// TwinCAT 3 PLC project Syn_Config
// Title: SynConfig
// Company: Syntegon Group
// ProjectVersion: 2.4.0.0
// Description: Parameter sets the RPP configurator writes and the application takes over (ADR 0017).
// ProgramVersion: 3.1.4026.28
// libraries:
//   Tc2_Standard,newest,Beckhoff Automation GmbH
//   SynVisu, * (Syntegon Group)
// project tree:
//   DUTs/ E_ConfigCommand.TcDUT, E_ConfigCommandResult.TcDUT, E_ConfigFieldType.TcDUT, E_ConfigResult.TcDUT, ST_ConfigBodyComponent.TcDUT, ST_ConfigBodyComponentParam.TcDUT, ST_ConfigBodyComponentSet.TcDUT, ST_ConfigCartesian.TcDUT, ST_ConfigCartesianParam.TcDUT, ST_ConfigCartesianSet.TcDUT, ST_ConfigCommand.TcDUT, ST_ConfigCommandStatus.TcDUT, ST_ConfigConveyor.TcDUT, ST_ConfigConveyorParam.TcDUT, ST_ConfigConveyorSet.TcDUT, ST_ConfigDelta.TcDUT, ST_ConfigDeltaParam.TcDUT, ST_ConfigDeltaSet.TcDUT, ST_ConfigMachine.TcDUT, ST_ConfigManifest.TcDUT, ST_ConfigManifestEntry.TcDUT, ST_ConfigRecipeField.TcDUT, ST_ConfigRecipeSet.TcDUT, ST_ConfigStaging.TcDUT, ST_ConfigStatus.TcDUT, ST_ConfigTopology.TcDUT, ST_ConfigTopologyKind.TcDUT, ST_ConfigTopologyLink.TcDUT, ST_ConfigTopologyLinks.TcDUT, ST_ConfigTopologyNode.TcDUT, ST_ConfigTopologyRole.TcDUT, ST_ConfigXtsGantry.TcDUT, ST_ConfigXtsGantryParam.TcDUT, ST_ConfigXtsGantrySet.TcDUT, ST_ConfigXtsLoop.TcDUT, ST_ConfigXtsLoopParam.TcDUT, ST_ConfigXtsLoopSet.TcDUT
//   GVLs/ CONFIG_GlobalConst.TcGVL, CONFIG_GlobalConst_Param.TcGVL
//   POUs/ _FB_ConfigBodyComponent.TcPOU, _FB_ConfigCartesian.TcPOU, _FB_ConfigComponent.TcPOU, _FB_ConfigConveyor.TcPOU, _FB_ConfigDelta.TcPOU, _FB_ConfigMachine.TcPOU, _FB_ConfigSensor.TcPOU, _FB_ConfigStation.TcPOU, _FB_ConfigTopology.TcPOU, _FB_ConfigVision.TcPOU, _FB_ConfigXtsGantry.TcPOU, _FB_ConfigXtsLoop.TcPOU, _FC_GetVersionSynConfig.TcPOU
// (motion and I/O tree: see PLC project syn_visu)
// real-time tasks:
//   TASK PlcTask: cycle T#10ms, priority 20, ADS port 350
//   TASK TestTask: cycle T#10ms, priority 21, ADS port 351

// ---- DUTs/E_ConfigCommand.TcDUT
{attribute 'qualified_only'}
{attribute 'strict'}
TYPE E_ConfigCommand :
(
	(* What a machine command asks the application (config protocol 3). Values are part of the gateway contract:
	   append, never renumber. *)
	NONE := 0,
	START := 1,
	STOP := 2,
	RESET := 3
) UINT;
END_TYPE

// ---- DUTs/E_ConfigCommandResult.TcDUT
{attribute 'qualified_only'}
{attribute 'strict'}
TYPE E_ConfigCommandResult :
(
	(* What the application made of the last machine command. Values are part of the gateway contract: append, never
	   renumber. *)
	NONE := 0,		// nothing asked since the PLC started
	ACCEPTED := 1,
	REJECTED := 2	// ST_ConfigCommandStatus.sMessage says why
) UINT;
END_TYPE

// ---- DUTs/E_ConfigFieldType.TcDUT
{attribute 'qualified_only'}
{attribute 'strict'}
TYPE E_ConfigFieldType :
(
	(* How a recipe field's value is kept (config protocol 3). Every value travels as LREAL. Values are part of the
	   gateway contract: append, never renumber. *)
	NUMBER := 0,	// any number within fMin..fMax
	INTEGER := 1,	// a whole number within fMin..fMax, e.g. picks per cycle
	SWITCH := 2,	// on or off: 1 or 0
	CHOICE := 3		// one of the named choices: 0..nChoiceCount-1
) UINT;
END_TYPE

// ---- DUTs/E_ConfigResult.TcDUT
{attribute 'qualified_only'}
{attribute 'strict'}
TYPE E_ConfigResult :
(
	(* What became of the last staged parameter set. Values are part of the gateway contract: append, never renumber. *)
	NONE := 0,		// nothing staged since the PLC started
	PENDING := 1,	// staged, waiting for the application to allow taking it over
	APPLIED := 2,	// taken over (or reset to the program values)
	REJECTED := 3	// not taken over; ST_ConfigStatus.sMessage says why
) UINT;
END_TYPE

// ---- DUTs/ST_ConfigBodyComponent.TcDUT
TYPE ST_ConfigBodyComponent :
STRUCT
	(* vo_Config of _FB_ConfigVision, _FB_ConfigSensor and _FB_ConfigStation: the gateway writes stStaging and
	   stStaged, reads stStatus and stActive. *)
	stStaging : ST_ConfigStaging;
	stStaged : ST_ConfigBodyComponentParam;
	stStatus : ST_ConfigStatus;
	stActive : ST_ConfigBodyComponentParam; // effective values: the active set while one is valid, else the program values
END_STRUCT
END_TYPE

// ---- DUTs/ST_ConfigBodyComponentParam.TcDUT
TYPE ST_ConfigBodyComponentParam :
STRUCT
	(* The parameter set of a component drawn from its bodies (vision system, product sensor, station): what the
	   configurator writes, never its bodies (hardware). Members as in SynVisu.ST_VisuDetectorConfig. *)
	stPose : SynVisu.ST_VisuPose; // MCS
	stOriginShift : SynVisu.ST_VisuPosition; // mm in the component's local frame
	nZoneCount : UINT;
	aZones : ARRAY[0..SynVisu.VISU_GlobalConst_Param.VISU_un_MAX_ZONES - 1] OF SynVisu.ST_VisuZone;
END_STRUCT
END_TYPE

// ---- DUTs/ST_ConfigBodyComponentSet.TcDUT
TYPE ST_ConfigBodyComponentSet :
STRUCT
	(* The active parameter set of a vision system, product sensor or station as the application keeps it, in a
	   VAR PERSISTENT variable passed to m_Cycle of _FB_ConfigVision, _FB_ConfigSensor or _FB_ConfigStation. *)
	bValid : BOOL; // FALSE: no set active, the program values apply
	nVersion : UDINT; // version of stParam
	nLastVersion : UDINT; // last version handed out; versions never repeat, also after a reset
	stParam : ST_ConfigBodyComponentParam;
END_STRUCT
END_TYPE

// ---- DUTs/ST_ConfigCartesian.TcDUT
TYPE ST_ConfigCartesian :
STRUCT
	(* vo_Config of _FB_ConfigCartesian: the gateway writes stStaging and stStaged, reads stStatus and stActive. *)
	stStaging : ST_ConfigStaging;
	stStaged : ST_ConfigCartesianParam;
	stStatus : ST_ConfigStatus;
	stActive : ST_ConfigCartesianParam; // effective values: the active set while one is valid, else the program values
END_STRUCT
END_TYPE

// ---- DUTs/ST_ConfigCartesianParam.TcDUT
TYPE ST_ConfigCartesianParam :
STRUCT
	(* A Cartesian robot's parameter set: what the configurator writes, never its axes, strokes or rail height
	   (hardware). Members as in SynVisu.ST_VisuCartesianConfig. *)
	stPose : SynVisu.ST_VisuPose; // MCS, axis origin X = Y = 0 with Z up
	stOriginShift : SynVisu.ST_VisuPosition; // mm in the robot's local frame
	nZoneCount : UINT;
	aZones : ARRAY[0..SynVisu.VISU_GlobalConst_Param.VISU_un_MAX_ZONES - 1] OF SynVisu.ST_VisuZone;
	nFingerCount : UINT; // gripper fingers with their flange offsets (config protocol 2, ADR 0018)
	aFingers : ARRAY[0..SynVisu.VISU_GlobalConst_Param.VISU_un_MAX_FINGERS - 1] OF SynVisu.ST_VisuFinger;
	stLimitArea : SynVisu.ST_VisuLimitArea; // bActive = FALSE: none
	stTcpLimitArea : SynVisu.ST_VisuLimitArea; // bActive = FALSE: none
END_STRUCT
END_TYPE

// ---- DUTs/ST_ConfigCartesianSet.TcDUT
TYPE ST_ConfigCartesianSet :
STRUCT
	(* A Cartesian robot's active parameter set as the application keeps it, in a VAR PERSISTENT variable passed to
	   _FB_ConfigCartesian.m_Cycle. *)
	bValid : BOOL; // FALSE: no set active, the program values apply
	nVersion : UDINT; // version of stParam
	nLastVersion : UDINT; // last version handed out; versions never repeat, also after a reset
	stParam : ST_ConfigCartesianParam;
END_STRUCT
END_TYPE

// ---- DUTs/ST_ConfigCommand.TcDUT
TYPE ST_ConfigCommand :
STRUCT
	(* A machine command, written by the gateway with bRequested last (config protocol 3). The machine FB clears
	   bRequested once the application answered it. *)
	nCommandId : UDINT; // chosen by the gateway; ST_ConfigCommandStatus.nHandledCommandId names it once answered
	eCommand : E_ConfigCommand;
	bRequested : BOOL; // TRUE: the command waits for the application's answer
END_STRUCT
END_TYPE

// ---- DUTs/ST_ConfigCommandStatus.TcDUT
TYPE ST_ConfigCommandStatus :
STRUCT
	nHandledCommandId : UDINT; // nCommandId of the last command the application answered
	eResult : E_ConfigCommandResult; // what the application made of it
	sMessage : STRING(80); // why it was rejected; empty otherwise
END_STRUCT
END_TYPE

// ---- DUTs/ST_ConfigConveyor.TcDUT
TYPE ST_ConfigConveyor :
STRUCT
	(* vo_Config of _FB_ConfigConveyor: the gateway writes stStaging and stStaged, reads stStatus and stActive. *)
	stStaging : ST_ConfigStaging;
	stStaged : ST_ConfigConveyorParam;
	stStatus : ST_ConfigStatus;
	stActive : ST_ConfigConveyorParam; // effective values: the active set while one is valid, else the program values
END_STRUCT
END_TYPE

// ---- DUTs/ST_ConfigConveyorParam.TcDUT
TYPE ST_ConfigConveyorParam :
STRUCT
	(* A conveyor's parameter set: what the configurator writes, never the belt's length or width (hardware).
	   Members as in SynVisu.ST_VisuConveyorConfig. *)
	stPose : SynVisu.ST_VisuPose; // MCS, belt start on the belt surface; local +X = conveying direction
	stOriginShift : SynVisu.ST_VisuPosition; // mm in the local frame from stPose: origin of the belt coordinates
	nProductTypeCount : UINT;
	aProductTypes : ARRAY[0..SynVisu.VISU_GlobalConst_Param.VISU_un_MAX_PRODUCT_TYPES - 1] OF SynVisu.ST_VisuProductType;
END_STRUCT
END_TYPE

// ---- DUTs/ST_ConfigConveyorSet.TcDUT
TYPE ST_ConfigConveyorSet :
STRUCT
	(* A conveyor's active parameter set as the application keeps it, in a VAR PERSISTENT variable passed to
	   _FB_ConfigConveyor.m_Cycle. *)
	bValid : BOOL; // FALSE: no set active, the program values apply
	nVersion : UDINT; // version of stParam
	nLastVersion : UDINT; // last version handed out; versions never repeat, also after a reset
	stParam : ST_ConfigConveyorParam;
END_STRUCT
END_TYPE

// ---- DUTs/ST_ConfigDelta.TcDUT
TYPE ST_ConfigDelta :
STRUCT
	(* vo_Config of _FB_ConfigDelta: the gateway writes stStaging and stStaged, reads stStatus and stActive. *)
	stStaging : ST_ConfigStaging;
	stStaged : ST_ConfigDeltaParam;
	stStatus : ST_ConfigStatus;
	stActive : ST_ConfigDeltaParam; // effective values: the active set while one is valid, else the program values
END_STRUCT
END_TYPE

// ---- DUTs/ST_ConfigDeltaParam.TcDUT
TYPE ST_ConfigDeltaParam :
STRUCT
	(* A Delta robot's parameter set: what the configurator writes, never its arm geometry (hardware).
	   Members as in SynVisu.ST_VisuDeltaConfig. *)
	stPose : SynVisu.ST_VisuPose; // MCS, base centre
	stOriginShift : SynVisu.ST_VisuPosition; // mm in the base's local frame
	nZoneCount : UINT;
	aZones : ARRAY[0..SynVisu.VISU_GlobalConst_Param.VISU_un_MAX_ZONES - 1] OF SynVisu.ST_VisuZone;
	nFingerCount : UINT; // gripper fingers with their flange offsets (config protocol 2, ADR 0018)
	aFingers : ARRAY[0..SynVisu.VISU_GlobalConst_Param.VISU_un_MAX_FINGERS - 1] OF SynVisu.ST_VisuFinger;
	stWorkingArea : SynVisu.ST_VisuWorkingArea;
	stLimitArea : SynVisu.ST_VisuLimitArea; // bActive = FALSE: none
	stTcpLimitArea : SynVisu.ST_VisuLimitArea; // bActive = FALSE: none
END_STRUCT
END_TYPE

// ---- DUTs/ST_ConfigDeltaSet.TcDUT
TYPE ST_ConfigDeltaSet :
STRUCT
	(* A Delta robot's active parameter set as the application keeps it, in a VAR PERSISTENT variable passed to
	   _FB_ConfigDelta.m_Cycle. *)
	bValid : BOOL; // FALSE: no set active, the program values apply
	nVersion : UDINT; // version of stParam
	nLastVersion : UDINT; // last version handed out; versions never repeat, also after a reset
	stParam : ST_ConfigDeltaParam;
END_STRUCT
END_TYPE

// ---- DUTs/ST_ConfigMachine.TcDUT
TYPE ST_ConfigMachine :
STRUCT
	(* vo_Config of _FB_ConfigMachine (config protocol 3, ADR 0022), listed in the config manifest with id 0 and type
	   NONE. The gateway reads the declared fields once, writes stStaging with aStaged (bStaged or bReset last) and
	   stCommand (bRequested last), and reads stStatus, aActive and stCommandStatus every cycle. Values are kept by
	   field index, every type as LREAL (SWITCH 0 / 1, INTEGER and CHOICE whole numbers). *)
	nFieldCount : UINT; // fields [0..nFieldCount-1] are declared
	aFields : ARRAY[0..CONFIG_GlobalConst_Param.CONFIG_un_MAX_RECIPE_FIELDS - 1] OF ST_ConfigRecipeField;
	stStaging : ST_ConfigStaging;
	aStaged : ARRAY[0..CONFIG_GlobalConst_Param.CONFIG_un_MAX_RECIPE_FIELDS - 1] OF LREAL; // the proposed recipe
	stStatus : ST_ConfigStatus;
	aActive : ARRAY[0..CONFIG_GlobalConst_Param.CONFIG_un_MAX_RECIPE_FIELDS - 1] OF LREAL; // effective values
	stCommand : ST_ConfigCommand;
	stCommandStatus : ST_ConfigCommandStatus;
END_STRUCT
END_TYPE

// ---- DUTs/ST_ConfigManifest.TcDUT
TYPE ST_ConfigManifest :
STRUCT
	(* Where the gateway finds the parameter FBs (ADR 0017). The application declares one instance at the symbol
	   GVL_Config.stManifest; every parameter FB registers itself with m_Register. *)
	nProtocolVersion : UINT := CONFIG_GlobalConst.CONFIG_un_PROTOCOL_VERSION;
	sLibraryVersion : STRING(15); // version of the Syn_Config library actually running, e.g. '1.0.0'
	nCount : UINT; // entries [0..nCount-1] are evaluated
	aEntries : ARRAY[0..CONFIG_GlobalConst_Param.CONFIG_un_MAX_MANIFEST_ENTRIES - 1] OF ST_ConfigManifestEntry;
END_STRUCT
END_TYPE

// ---- DUTs/ST_ConfigManifestEntry.TcDUT
TYPE ST_ConfigManifestEntry :
STRUCT
	nId : UDINT; // manifest id of the Syn_Visu component the parameter FB is for
	eType : SynVisu.E_VisuComponentType; // type of that component
	sPath : STRING(255); // symbol path of the parameter FB's vo_Config, e.g. 'P_Line.fb_InfeedParam.vo_Config'
END_STRUCT
END_TYPE

// ---- DUTs/ST_ConfigRecipeField.TcDUT
TYPE ST_ConfigRecipeField :
STRUCT
	(* One field of the machine's recipe as the application declares it with _FB_ConfigMachine.m_DeclareField
	   (config protocol 3, ADR 0022), m_SetText and m_SetVisibleWhen (config protocol 4, #49). The gateway reads the
	   declarations once at discovery. *)
	sName : STRING(31); // unique in the recipe, e.g. 'BeltSpeed'
	nGroup : UDINT; // manifest id of the Syn_Visu component the field belongs to, 0 = the whole machine
	eType : E_ConfigFieldType;
	sUnit : STRING(15); // e.g. 'mm/s', '' = none
	fMin : LREAL; // smallest value of a NUMBER or INTEGER field
	fMax : LREAL; // largest value of a NUMBER or INTEGER field
	fProgramValue : LREAL; // the application's own value, which applies while no recipe is active
	nChoiceCount : UINT; // named values of a CHOICE field
	aChoices : ARRAY[0..CONFIG_GlobalConst_Param.CONFIG_un_MAX_CHOICES - 1] OF STRING(31); // their names, from value 0
	sLabel : STRING(40); // what the Simulator calls the field, '' = its name put into words
	sDescription : STRING(160); // what the field is for, shown in its tooltip, '' = none
	nVisibleField : UINT; // the field (from 1) it applies only with, 0 = always
	nVisibleValue : DINT; // the value nVisibleField must have: a SWITCH's 0 / 1, a CHOICE's number, a whole number
END_STRUCT
END_TYPE

// ---- DUTs/ST_ConfigRecipeSet.TcDUT
TYPE ST_ConfigRecipeSet :
STRUCT
	(* The machine's active recipe as the application keeps it, in a VAR PERSISTENT variable passed to
	   _FB_ConfigMachine.m_Cycle. Values by field index: keep the fields' order, add new ones at the end. *)
	bValid : BOOL; // FALSE: no recipe active, the program values apply
	nVersion : UDINT; // version of aValues
	nLastVersion : UDINT; // last version handed out; versions never repeat, also after a reset
	aValues : ARRAY[0..CONFIG_GlobalConst_Param.CONFIG_un_MAX_RECIPE_FIELDS - 1] OF LREAL;
END_STRUCT
END_TYPE

// ---- DUTs/ST_ConfigStaging.TcDUT
TYPE ST_ConfigStaging :
STRUCT
	(* Written by the gateway in one ADS sum-write, bStaged or bReset last, so a set is never seen staged half
	   written (ADR 0017). The parameter FB clears bStaged and bReset once it handled them. *)
	nBaseVersion : UDINT; // active version the staged set is based on; another active version rejects it
	nStageId : UDINT; // chosen by the gateway; ST_ConfigStatus.nHandledStageId names it once handled
	bReset : BOOL; // TRUE: make the active set invalid, the program values apply again
	bStaged : BOOL; // TRUE: stStaged is complete and waits to be taken over
END_STRUCT
END_TYPE

// ---- DUTs/ST_ConfigStatus.TcDUT
TYPE ST_ConfigStatus :
STRUCT
	nActiveVersion : UDINT; // version of the active set; 0 while the program values apply
	nHandledStageId : UDINT; // nStageId of the last staging handled (taken over, rejected or reset)
	eResult : E_ConfigResult; // what became of it
	sMessage : STRING(80); // why it was rejected; empty otherwise
END_STRUCT
END_TYPE

// ---- DUTs/ST_ConfigTopology.TcDUT
TYPE ST_ConfigTopology :
STRUCT
	(* vo_Config of _FB_ConfigTopology (config protocol 5, ADR 0023), listed in the config manifest with id 0 and type
	   NONE like the machine FB; the gateway tells them apart by this type. It reads the declaration once at discovery
	   and stActive every cycle. *)
	nKindCount : UINT; // kinds [0..nKindCount-1] are declared
	aKinds : ARRAY[0..CONFIG_GlobalConst_Param.CONFIG_un_MAX_TOPOLOGY_KINDS - 1] OF ST_ConfigTopologyKind;
	nRoleCount : UINT; // roles [0..nRoleCount-1] are declared
	aRoles : ARRAY[0..CONFIG_GlobalConst_Param.CONFIG_un_MAX_TOPOLOGY_ROLES - 1] OF ST_ConfigTopologyRole;
	nNodeCount : UINT; // nodes [0..nNodeCount-1] are declared
	aNodes : ARRAY[0..CONFIG_GlobalConst_Param.CONFIG_un_MAX_TOPOLOGY_NODES - 1] OF ST_ConfigTopologyNode;
	nRootNode : DINT; // id of the root node, which has no parent; 0 = none set
	stActive : ST_ConfigTopologyLinks; // the links in effect: the application's program values
END_STRUCT
END_TYPE

// ---- DUTs/ST_ConfigTopologyKind.TcDUT
TYPE ST_ConfigTopologyKind :
STRUCT
	(* A kind of topology node as the application declares it with _FB_ConfigTopology.m_DeclareKind (config protocol 5,
	   ADR 0023), referred to by its number from 1. *)
	sName : STRING(31); // unique in the topology, e.g. 'PPH'
	nParentKinds : DWORD; // bit k - 1 set: a node of kind k may be the parent of a node of this kind (m_AllowParent)
END_STRUCT
END_TYPE

// ---- DUTs/ST_ConfigTopologyLink.TcDUT
TYPE ST_ConfigTopologyLink :
STRUCT
	(* One link of a topology (config protocol 5, ADR 0023): node nNode points to node nTarget in role nRole. *)
	nNode : DINT; // id of the node that holds the link
	nRole : UINT; // its role, from 1; 0 = nTarget is the node's parent
	nTarget : DINT; // id of the node it points to
END_STRUCT
END_TYPE

// ---- DUTs/ST_ConfigTopologyLinks.TcDUT
TYPE ST_ConfigTopologyLinks :
STRUCT
	(* The links of a topology, its parents included (config protocol 5, ADR 0023). *)
	nLinkCount : UINT; // links [0..nLinkCount-1] are set
	aLinks : ARRAY[0..CONFIG_GlobalConst_Param.CONFIG_un_MAX_TOPOLOGY_LINKS - 1] OF ST_ConfigTopologyLink;
END_STRUCT
END_TYPE

// ---- DUTs/ST_ConfigTopologyNode.TcDUT
TYPE ST_ConfigTopologyNode :
STRUCT
	(* One topology node of the full build-out as the application declares it with _FB_ConfigTopology.m_DeclareNode and
	   m_AddComponent (config protocol 5, ADR 0023). *)
	nId : DINT; // the application's id, unique in the topology, e.g. its context id
	sName : STRING(31); // e.g. 'PPH1'
	nKind : UINT; // its kind, from 1
	nComponentCount : UINT; // Syn_Visu components the node stands for
	aComponents : ARRAY[0..CONFIG_GlobalConst_Param.CONFIG_un_MAX_NODE_COMPONENTS - 1] OF UDINT; // their manifest ids
END_STRUCT
END_TYPE

// ---- DUTs/ST_ConfigTopologyRole.TcDUT
TYPE ST_ConfigTopologyRole :
STRUCT
	(* What a topology link means, as the application declares it with _FB_ConfigTopology.m_DeclareRole (config
	   protocol 5, ADR 0023), referred to by its number from 1; role 0 is the parent. *)
	sName : STRING(31); // unique in the topology, e.g. 'Infeed1'
	nHolderKind : UINT; // the kind (from 1) of node that holds the role
	nTargetKinds : DWORD; // bit k - 1 set: a link in this role may point to a node of kind k (m_AllowTarget)
	bRequired : BOOL; // a node in use of the holder kind must have a link in this role
END_STRUCT
END_TYPE

// ---- DUTs/ST_ConfigXtsGantry.TcDUT
TYPE ST_ConfigXtsGantry :
STRUCT
	(* vo_Config of _FB_ConfigXtsGantry: the gateway writes stStaging and stStaged, reads stStatus and stActive. *)
	stStaging : ST_ConfigStaging;
	stStaged : ST_ConfigXtsGantryParam;
	stStatus : ST_ConfigStatus;
	stActive : ST_ConfigXtsGantryParam; // effective values: the active set while one is valid, else the program values
END_STRUCT
END_TYPE

// ---- DUTs/ST_ConfigXtsGantryParam.TcDUT
TYPE ST_ConfigXtsGantryParam :
STRUCT
	(* An XTS gantry's parameter set: what the configurator writes, never its strokes, tool offsets or mover size
	   (hardware). Members as in SynVisu.ST_VisuXtsGantryConfig. *)
	stPose : SynVisu.ST_VisuPose; // MCS, track start on top of the movers with Z = 0
	stOriginShift : SynVisu.ST_VisuPosition; // mm in the track's local frame
	nModuleCount : UINT;
	aModules : ARRAY[0..SynVisu.VISU_GlobalConst_Param.VISU_un_MAX_MODULES - 1] OF SynVisu.ST_VisuTrackModule;
	nZoneCount : UINT;
	aZones : ARRAY[0..SynVisu.VISU_GlobalConst_Param.VISU_un_MAX_ZONES - 1] OF SynVisu.ST_VisuZone;
	nFingerCount : UINT; // gripper fingers of every mover, with their flange offsets (config protocol 2, ADR 0018)
	aFingers : ARRAY[0..SynVisu.VISU_GlobalConst_Param.VISU_un_MAX_FINGERS - 1] OF SynVisu.ST_VisuFinger;
	stLimitArea : SynVisu.ST_VisuLimitArea; // bActive = FALSE: none
	stTcpLimitArea : SynVisu.ST_VisuLimitArea; // bActive = FALSE: none
END_STRUCT
END_TYPE

// ---- DUTs/ST_ConfigXtsGantrySet.TcDUT
TYPE ST_ConfigXtsGantrySet :
STRUCT
	(* An XTS gantry's active parameter set as the application keeps it, in a VAR PERSISTENT variable passed to
	   _FB_ConfigXtsGantry.m_Cycle. *)
	bValid : BOOL; // FALSE: no set active, the program values apply
	nVersion : UDINT; // version of stParam
	nLastVersion : UDINT; // last version handed out; versions never repeat, also after a reset
	stParam : ST_ConfigXtsGantryParam;
END_STRUCT
END_TYPE

// ---- DUTs/ST_ConfigXtsLoop.TcDUT
TYPE ST_ConfigXtsLoop :
STRUCT
	(* vo_Config of _FB_ConfigXtsLoop: the gateway writes stStaging and stStaged, reads stStatus and stActive. *)
	stStaging : ST_ConfigStaging;
	stStaged : ST_ConfigXtsLoopParam;
	stStatus : ST_ConfigStatus;
	stActive : ST_ConfigXtsLoopParam; // effective values: the active set while one is valid, else the program values
END_STRUCT
END_TYPE

// ---- DUTs/ST_ConfigXtsLoopParam.TcDUT
TYPE ST_ConfigXtsLoopParam :
STRUCT
	(* An XTS loop's parameter set: what the configurator writes, never its tool offset or mover size (hardware).
	   Members as in SynVisu.ST_VisuXtsLoopConfig. *)
	stPose : SynVisu.ST_VisuPose; // MCS, start of module 1
	stOriginShift : SynVisu.ST_VisuPosition; // mm in the loop's local frame
	nModuleCount : UINT;
	aModules : ARRAY[0..SynVisu.VISU_GlobalConst_Param.VISU_un_MAX_MODULES - 1] OF SynVisu.ST_VisuTrackModule;
	nZoneCount : UINT;
	aZones : ARRAY[0..SynVisu.VISU_GlobalConst_Param.VISU_un_MAX_ZONES - 1] OF SynVisu.ST_VisuZone;
	nFingerCount : UINT; // gripper fingers of every mover, with their flange offsets (config protocol 2, ADR 0018)
	aFingers : ARRAY[0..SynVisu.VISU_GlobalConst_Param.VISU_un_MAX_FINGERS - 1] OF SynVisu.ST_VisuFinger;
END_STRUCT
END_TYPE

// ---- DUTs/ST_ConfigXtsLoopSet.TcDUT
TYPE ST_ConfigXtsLoopSet :
STRUCT
	(* An XTS loop's active parameter set as the application keeps it, in a VAR PERSISTENT variable passed to
	   _FB_ConfigXtsLoop.m_Cycle. *)
	bValid : BOOL; // FALSE: no set active, the program values apply
	nVersion : UDINT; // version of stParam
	nLastVersion : UDINT; // last version handed out; versions never repeat, also after a reset
	stParam : ST_ConfigXtsLoopParam;
END_STRUCT
END_TYPE

// ---- GVLs/CONFIG_GlobalConst.TcGVL
(****************************************************************************************************<br>
© Syntegon Group.<br>
All rights reserved, also regarding any disposal, exploitation, reproduction, editing, distribution,<br>
as well as in the event of applications for industrial property rights.<br>
*****************************************************************************************************<br>
DESCRIPTION:<br>
Global constants of the Syn_Config library.<br>
****************************************************************************************************)
{attribute 'qualified_only'}
VAR_GLOBAL CONSTANT
	(* Version of the Syn_Config <-> gateway contract (ADR 0017). The gateway writes nothing to a PLC whose config
	   manifest reports a version it does not know (it knows 2 to 5). Bump together with CONFIG_PROTOCOL_VERSION in
	   the gateway.
	   1: conveyor (pose, origin shift, product types) and Delta (pose, origin shift, zones, working, limit and
	      TCP limit area); since library 1.1.0 also XTS gantry, XTS loop, Cartesian, vision, sensor and station
	      (new parameter FBs only: no change for a gateway or an application of 1.0.0).
	   2: gripper fingers with their flange offsets (nFingerCount, aFingers) in the parameter sets of the Delta,
	      the XTS gantry and loop and the Cartesian robot (library 2.0.0, ADR 0018).
	   3: the machine FB _FB_ConfigMachine (id 0, type NONE in the manifest): recipe fields the application declares,
	      their staging, and machine commands (library 2.1.0, ADR 0022). A PLC of version 2 still gets its parameter
	      sets written, but no recipe and no commands.
	   4: a recipe field's label, description and visibility condition (sLabel, sDescription, nVisibleField,
	      nVisibleValue; library 2.2.0, #49). A gateway reads the fields of version 3 without them.
	   5: the topology FB _FB_ConfigTopology (id 0, type NONE like the machine FB, told apart by the type of its
	      vo_Config): the application's topology nodes, roles and links (library 2.4.0, ADR 0023). *)
	CONFIG_un_PROTOCOL_VERSION			: UINT := 5;
	(* Version of this library (config manifest sLibraryVersion). Bump together with _FC_GetVersionSynConfig and the
	   project version. *)
	CONFIG_str_LIBRARY_VERSION			: STRING(15) := '2.4.0';
END_VAR

// ---- GVLs/CONFIG_GlobalConst_Param.TcGVL
(****************************************************************************************************<br>
© Syntegon Group.<br>
All rights reserved, also regarding any disposal, exploitation, reproduction, editing, distribution,<br>
as well as in the event of applications for industrial property rights.<br>
*****************************************************************************************************<br>
DESCRIPTION:<br>
Library parameters of Syn_Config: array sizes of the interface structures. The lists of a parameter set have the
sizes of Syn_Visu's (VISU_GlobalConst_Param), so every set fits the visualisation it is passed on to.<br>
****************************************************************************************************)
{attribute 'qualified_only'}
VAR_GLOBAL CONSTANT
	CONFIG_un_MAX_MANIFEST_ENTRIES		: UINT := 32;	// [-] parameter FBs in the config manifest
	CONFIG_un_MAX_RECIPE_FIELDS			: UINT := 64;	// [-] fields of the machine's recipe (_FB_ConfigMachine)
	CONFIG_un_MAX_CHOICES				: UINT := 8;	// [-] named values of a CHOICE recipe field
	CONFIG_un_MAX_TOPOLOGY_KINDS		: UINT := 16;	// [-] kinds of topology node (_FB_ConfigTopology), at most 32
	CONFIG_un_MAX_TOPOLOGY_ROLES		: UINT := 16;	// [-] roles a topology link may have
	CONFIG_un_MAX_TOPOLOGY_NODES		: UINT := 64;	// [-] topology nodes of the full build-out
	CONFIG_un_MAX_TOPOLOGY_LINKS		: UINT := 128;	// [-] links of a topology, its parents included
	CONFIG_un_MAX_NODE_COMPONENTS		: UINT := 4;	// [-] Syn_Visu components one topology node stands for
END_VAR

// ---- POUs/_FB_ConfigMachine.TcPOU
(****************************************************************************************************<br>
© Syntegon Group.<br>
All rights reserved, also regarding any disposal, exploitation, reproduction, editing, distribution,<br>
as well as in the event of applications for industrial property rights.<br>
*****************************************************************************************************<br>
DESCRIPTION:<br>
The machine as a whole (config protocol 3, ADR 0022): the recipe fields the application declares (process values<br>
such as belt speed, picks per cycle, the product pattern), their staging by the Simulator with the mechanism of the<br>
parameter sets, and the machine commands Start, Stop and Reset the application answers. One per application,<br>
listed in the config manifest with id 0. Typical cycle:<br>
  fb_Machine.m_Register(vio_Manifest := GVL_Config.stManifest, vi_udn_Id := 0);<br>
  fb_Machine.m_DeclareField(vi_un_Field := 1, vi_str_Name := 'BeltSpeed', vi_udn_Group := fb_Infeed.m_Id(),<br>
    vi_e_Type := E_ConfigFieldType.NUMBER, vi_str_Unit := 'mm/s', vi_lr_Min := 0, vi_lr_Max := 500,<br>
    vi_lr_ProgramValue := 150);<br>
  fb_Machine.m_SetText(vi_un_Field := 1, vi_str_Label := 'Belt speed', vi_str_Description := 'Speed of the infeed');<br>
  fb_Machine.m_SetVisibleWhen(vi_un_Field := 3, vi_un_OnField := 2, vi_dn_Value := 0);  // field 3 only with 2 = 0<br>
  fb_Machine.m_Cycle(vio_Set := RecipeSet, vi_b_ApplyAllowed := b_Stopped);<br>
  lr_BeltSpeed := fb_Machine.m_Value(vi_un_Field := 1);<br>
  CASE fb_Machine.m_Command() OF E_ConfigCommand.START: ...<br>
    fb_Machine.m_AnswerCommand(vi_b_Accepted := TRUE, vi_str_Reason := ''); END_CASE<br>
RecipeSet is the application's VAR PERSISTENT ST_ConfigRecipeSet.<br>
*****************************************************************************************************<br>
OUTPUT VALUES:<br>
vo_Config is the contract structure the gateway reads and writes at the path in the config manifest.<br>
*****************************************************************************************************<br>
LIMITS:<br>
CONFIG_un_MAX_RECIPE_FIELDS fields, CONFIG_un_MAX_CHOICES choices each. The gateway reads the declarations when<br>
it discovers the PLC: declare every field from the start and keep their order.<br>
*****************************************************************************************************<br>
VERSION         ¦ DATE       ¦ NAME      ¦ CHANGE<br>
Syn_Config 2.1.0 ¦ 2026-11-14 ¦ J.Willner ¦ Created: recipe fields and machine commands (protocol 3)<br>
Syn_Config 2.2.0 ¦ 2026-11-14 ¦ J.Willner ¦ m_SetText, m_SetVisibleWhen (protocol 4, #49)<br>
Syn_Config 2.3.0 ¦ 2026-11-14 ¦ J.Willner ¦ m_Cycle through m_HandleStaging<br>
****************************************************************************************************)
FUNCTION_BLOCK _FB_ConfigMachine EXTENDS _FB_ConfigComponent
VAR_OUTPUT
	vo_Config							: ST_ConfigMachine;	// contract structure of the gateway
END_VAR

(****************************************************************************************************<br>
© Syntegon Group.<br>
All rights reserved, also regarding any disposal, exploitation, reproduction, editing, distribution,<br>
as well as in the event of applications for industrial property rights.<br>
*****************************************************************************************************<br>
DESCRIPTION:<br>
Answers the waiting machine command: accepted, or rejected with the reason the Simulator shows. The command no<br>
longer waits afterwards.<br>
*****************************************************************************************************<br>
OUTPUT VALUES:<br>
FALSE while no command waits.<br>
****************************************************************************************************)
METHOD m_AnswerCommand : BOOL
VAR_INPUT
	vi_b_Accepted						: BOOL;	// TRUE: the application carries the command out
	vi_str_Reason						: STRING(80);	// why it is rejected, '' when accepted
END_VAR
m_AnswerCommand := vo_Config.stCommand.bRequested;
IF NOT m_AnswerCommand THEN
	RETURN;
END_IF
vo_Config.stCommandStatus.nHandledCommandId := vo_Config.stCommand.nCommandId;
vo_Config.stCommandStatus.eResult := SEL(vi_b_Accepted, E_ConfigCommandResult.REJECTED, E_ConfigCommandResult.ACCEPTED);
vo_Config.stCommandStatus.sMessage := SEL(vi_b_Accepted, vi_str_Reason, '');
vo_Config.stCommand.bRequested := FALSE;
END_METHOD

(****************************************************************************************************<br>
© Syntegon Group.<br>
All rights reserved, also regarding any disposal, exploitation, reproduction, editing, distribution,<br>
as well as in the event of applications for industrial property rights.<br>
*****************************************************************************************************<br>
DESCRIPTION:<br>
The machine command waiting for the application's answer (START, STOP, RESET); NONE while none waits. Answer it<br>
with m_AnswerCommand: the application alone decides whether it is carried out.<br>
****************************************************************************************************)
METHOD m_Command : E_ConfigCommand
IF vo_Config.stCommand.bRequested THEN
	m_Command := vo_Config.stCommand.eCommand;
ELSE
	m_Command := E_ConfigCommand.NONE;
END_IF
END_METHOD

(****************************************************************************************************<br>
© Syntegon Group.<br>
All rights reserved, also regarding any disposal, exploitation, reproduction, editing, distribution,<br>
as well as in the event of applications for industrial property rights.<br>
*****************************************************************************************************<br>
DESCRIPTION:<br>
Every cycle, after the fields are declared: handles a staged recipe or a reset (a recipe only while<br>
vi_b_ApplyAllowed), keeps the active recipe in vio_Set and gives the effective values in vo_Config.aActive: the<br>
active recipe while one is valid, else the fields' program values.<br>
*****************************************************************************************************<br>
OUTPUT VALUES:<br>
TRUE in the cycle a recipe was taken over or reset.<br>
****************************************************************************************************)
METHOD m_Cycle : BOOL
VAR_IN_OUT
	vio_Set								: ST_ConfigRecipeSet;	// the application's VAR PERSISTENT active recipe
END_VAR
VAR_INPUT
	vi_b_ApplyAllowed					: BOOL;	// [-] a staged recipe may be taken over now, e.g. while the machine stands
END_VAR
VAR
	b_TempTakeOver						: BOOL;	// the staged recipe was taken over: copy it
	un_TempIndex						: UINT;
END_VAR
m_Cycle := m_HandleStaging(vio_Staging := vo_Config.stStaging, vio_Status := vo_Config.stStatus, vio_b_Valid := vio_Set.bValid,
	vio_udn_Version := vio_Set.nVersion, vio_udn_LastVersion := vio_Set.nLastVersion, vi_b_ApplyAllowed := vi_b_ApplyAllowed,
	vo_b_TakeOver => b_TempTakeOver);
IF b_TempTakeOver THEN
	vio_Set.aValues := vo_Config.aStaged;
END_IF


(****************************************************************************************************
EFFECTIVE VALUES
****************************************************************************************************)
un_TempIndex := 0;
WHILE un_TempIndex < vo_Config.nFieldCount AND un_TempIndex < CONFIG_GlobalConst_Param.CONFIG_un_MAX_RECIPE_FIELDS DO
	vo_Config.aActive[un_TempIndex] := SEL(vio_Set.bValid, vo_Config.aFields[un_TempIndex].fProgramValue,
		vio_Set.aValues[un_TempIndex]);
	un_TempIndex := un_TempIndex + 1;
END_WHILE
END_METHOD

(****************************************************************************************************<br>
© Syntegon Group.<br>
All rights reserved, also regarding any disposal, exploitation, reproduction, editing, distribution,<br>
as well as in the event of applications for industrial property rights.<br>
*****************************************************************************************************<br>
DESCRIPTION:<br>
Declares recipe field vi_un_Field (1..CONFIG_un_MAX_RECIPE_FIELDS): its name, the component it belongs to, how its<br>
value is kept, its unit, range and the program value that applies while no recipe is active. Fields are listed up<br>
to the highest one declared. Idempotent: call it every cycle, before m_Cycle. A CHOICE field's values are named with<br>
m_SetChoice and range from 0; its vi_lr_Min and vi_lr_Max are not used, nor a SWITCH's.<br>
*****************************************************************************************************<br>
OUTPUT VALUES:<br>
FALSE for vi_un_Field = 0 or above CONFIG_un_MAX_RECIPE_FIELDS.<br>
****************************************************************************************************)
METHOD m_DeclareField : BOOL
VAR_INPUT
	vi_un_Field							: UINT;	// [-] 1..CONFIG_un_MAX_RECIPE_FIELDS
	vi_str_Name							: STRING(31);	// unique in the recipe, e.g. 'BeltSpeed'
	vi_udn_Group						: UDINT;	// [-] manifest id of the Syn_Visu component, 0 = the whole machine
	vi_e_Type							: E_ConfigFieldType;
	vi_str_Unit							: STRING(15);	// e.g. 'mm/s', '' = none
	vi_lr_Min							: LREAL;	// smallest value of a NUMBER or INTEGER field
	vi_lr_Max							: LREAL;	// largest value of a NUMBER or INTEGER field
	vi_lr_ProgramValue					: LREAL;	// the application's own value; a SWITCH: 1 = on
END_VAR
m_DeclareField := vi_un_Field > 0 AND vi_un_Field <= CONFIG_GlobalConst_Param.CONFIG_un_MAX_RECIPE_FIELDS;
IF NOT m_DeclareField THEN
	RETURN;
END_IF
vo_Config.aFields[vi_un_Field - 1].sName := vi_str_Name;
vo_Config.aFields[vi_un_Field - 1].nGroup := vi_udn_Group;
vo_Config.aFields[vi_un_Field - 1].eType := vi_e_Type;
vo_Config.aFields[vi_un_Field - 1].sUnit := vi_str_Unit;
vo_Config.aFields[vi_un_Field - 1].fMin := vi_lr_Min;
vo_Config.aFields[vi_un_Field - 1].fMax := vi_lr_Max;
vo_Config.aFields[vi_un_Field - 1].fProgramValue := vi_lr_ProgramValue;
IF vi_un_Field > vo_Config.nFieldCount THEN
	vo_Config.nFieldCount := vi_un_Field;
END_IF
END_METHOD

(****************************************************************************************************<br>
© Syntegon Group.<br>
All rights reserved, also regarding any disposal, exploitation, reproduction, editing, distribution,<br>
as well as in the event of applications for industrial property rights.<br>
*****************************************************************************************************<br>
DESCRIPTION:<br>
Effective value of an INTEGER or CHOICE recipe field as a whole number (see m_Value).<br>
****************************************************************************************************)
METHOD m_Integer : DINT
VAR_INPUT
	vi_un_Field							: UINT;	// [-] 1..the field count
END_VAR
m_Integer := LREAL_TO_DINT(m_Value(vi_un_Field := vi_un_Field));
END_METHOD

(****************************************************************************************************<br>
© Syntegon Group.<br>
All rights reserved, also regarding any disposal, exploitation, reproduction, editing, distribution,<br>
as well as in the event of applications for industrial property rights.<br>
*****************************************************************************************************<br>
DESCRIPTION:<br>
Why the staged recipe cannot be taken over; '' when it can: a value outside its field's range (NUMBER, INTEGER),<br>
not one of its choices (CHOICE), not a whole number (INTEGER, CHOICE) or not 0 or 1 (SWITCH).<br>
****************************************************************************************************)
METHOD PROTECTED m_InvalidStaged : STRING(80)
VAR
	un_TempIndex						: UINT;
	lr_TempValue						: LREAL;
	lr_TempMin							: LREAL;
	lr_TempMax							: LREAL;
END_VAR
m_InvalidStaged := '';
un_TempIndex := 0;
WHILE un_TempIndex < vo_Config.nFieldCount AND un_TempIndex < CONFIG_GlobalConst_Param.CONFIG_un_MAX_RECIPE_FIELDS DO
	lr_TempValue := vo_Config.aStaged[un_TempIndex];
	CASE vo_Config.aFields[un_TempIndex].eType OF
		E_ConfigFieldType.SWITCH:
			lr_TempMin := 0;
			lr_TempMax := 1;
		E_ConfigFieldType.CHOICE:
			lr_TempMin := 0;
			lr_TempMax := UINT_TO_LREAL(vo_Config.aFields[un_TempIndex].nChoiceCount) - 1;
	ELSE
		lr_TempMin := vo_Config.aFields[un_TempIndex].fMin;
		lr_TempMax := vo_Config.aFields[un_TempIndex].fMax;
	END_CASE
	(* The range first: only a value in range is turned into a whole number. NaN equals nothing, not even itself. *)
	IF lr_TempValue <> lr_TempValue OR lr_TempValue < lr_TempMin OR lr_TempValue > lr_TempMax THEN
		m_InvalidStaged := CONCAT(CONCAT('Field ', vo_Config.aFields[un_TempIndex].sName), CONCAT(': ', CONCAT(LREAL_TO_STRING(lr_TempValue),
			CONCAT(' is outside ', CONCAT(LREAL_TO_STRING(lr_TempMin), CONCAT(' to ', LREAL_TO_STRING(lr_TempMax)))))));
		RETURN;
	END_IF
	IF vo_Config.aFields[un_TempIndex].eType <> E_ConfigFieldType.NUMBER
		AND LINT_TO_LREAL(LREAL_TO_LINT(lr_TempValue)) <> lr_TempValue
	THEN
		m_InvalidStaged := CONCAT(CONCAT('Field ', vo_Config.aFields[un_TempIndex].sName), CONCAT(': ',
			CONCAT(LREAL_TO_STRING(lr_TempValue), ' is not a value of its type')));
		RETURN;
	END_IF
	un_TempIndex := un_TempIndex + 1;
END_WHILE
END_METHOD

(****************************************************************************************************<br>
© Syntegon Group.<br>
All rights reserved, also regarding any disposal, exploitation, reproduction, editing, distribution,<br>
as well as in the event of applications for industrial property rights.<br>
*****************************************************************************************************<br>
DESCRIPTION:<br>
Names value vi_un_Value (0..CONFIG_un_MAX_CHOICES-1) of the CHOICE field vi_un_Field, e.g. 0 = 'Lanes'. The field<br>
has as many choices as the highest value named plus one. Idempotent: call it every cycle with m_DeclareField.<br>
*****************************************************************************************************<br>
OUTPUT VALUES:<br>
FALSE for a field not declared or a value above CONFIG_un_MAX_CHOICES - 1.<br>
****************************************************************************************************)
METHOD m_SetChoice : BOOL
VAR_INPUT
	vi_un_Field							: UINT;	// [-] the field, 1..its count
	vi_un_Value							: UINT;	// [-] the value it names, from 0
	vi_str_Text							: STRING(31);	// e.g. 'Lanes'
END_VAR
m_SetChoice := vi_un_Field > 0 AND vi_un_Field <= vo_Config.nFieldCount
	AND vi_un_Value < CONFIG_GlobalConst_Param.CONFIG_un_MAX_CHOICES;
IF NOT m_SetChoice THEN
	RETURN;
END_IF
vo_Config.aFields[vi_un_Field - 1].aChoices[vi_un_Value] := vi_str_Text;
IF vi_un_Value >= vo_Config.aFields[vi_un_Field - 1].nChoiceCount THEN
	vo_Config.aFields[vi_un_Field - 1].nChoiceCount := vi_un_Value + 1;
END_IF
END_METHOD

(****************************************************************************************************<br>
© Syntegon Group.<br>
All rights reserved, also regarding any disposal, exploitation, reproduction, editing, distribution,<br>
as well as in the event of applications for industrial property rights.<br>
*****************************************************************************************************<br>
DESCRIPTION:<br>
Gives the declared field vi_un_Field the label the Simulator shows instead of its name put into words, and a<br>
description of what it is for, shown in the field's tooltip (config protocol 4, #49). Free text in the operators'<br>
language; the name stays the field's key. Idempotent: call it every cycle with m_DeclareField.<br>
*****************************************************************************************************<br>
OUTPUT VALUES:<br>
FALSE for a field not declared.<br>
****************************************************************************************************)
METHOD m_SetText : BOOL
VAR_INPUT
	vi_un_Field							: UINT;	// [-] the field, 1..its count
	vi_str_Label						: STRING(40);	// e.g. 'Belt speed', '' = the name put into words
	vi_str_Description					: STRING(160);	// what the field is for, '' = none
END_VAR
m_SetText := vi_un_Field > 0 AND vi_un_Field <= vo_Config.nFieldCount;
IF NOT m_SetText THEN
	RETURN;
END_IF
vo_Config.aFields[vi_un_Field - 1].sLabel := vi_str_Label;
vo_Config.aFields[vi_un_Field - 1].sDescription := vi_str_Description;
END_METHOD

(****************************************************************************************************<br>
© Syntegon Group.<br>
All rights reserved, also regarding any disposal, exploitation, reproduction, editing, distribution,<br>
as well as in the event of applications for industrial property rights.<br>
*****************************************************************************************************<br>
DESCRIPTION:<br>
Shows the declared field vi_un_Field in the Simulator only while field vi_un_OnField has the value vi_dn_Value<br>
(config protocol 4, #49), e.g. a lane count only while the pattern is Lanes. vi_un_OnField must be a SWITCH (0 / 1),<br>
CHOICE or INTEGER field and may belong to another group; a field depending on a hidden one is hidden too. A hidden<br>
field keeps its value and is written with the recipe. vi_un_OnField = 0 shows the field always. The gateway reports<br>
a condition on a NUMBER field, on the field itself, on a field not declared, on a value that field can never have<br>
or in a ring as a discovery error and shows that field always. Idempotent: call it every cycle with m_DeclareField.<br>
*****************************************************************************************************<br>
OUTPUT VALUES:<br>
FALSE for a field not declared.<br>
****************************************************************************************************)
METHOD m_SetVisibleWhen : BOOL
VAR_INPUT
	vi_un_Field							: UINT;	// [-] the field shown on condition, 1..its count
	vi_un_OnField						: UINT;	// [-] the field the condition reads, 0 = always shown
	vi_dn_Value							: DINT;	// [-] the value vi_un_OnField must have
END_VAR
m_SetVisibleWhen := vi_un_Field > 0 AND vi_un_Field <= vo_Config.nFieldCount;
IF NOT m_SetVisibleWhen THEN
	RETURN;
END_IF
vo_Config.aFields[vi_un_Field - 1].nVisibleField := vi_un_OnField;
vo_Config.aFields[vi_un_Field - 1].nVisibleValue := vi_dn_Value;
END_METHOD

(****************************************************************************************************<br>
© Syntegon Group.<br>
All rights reserved, also regarding any disposal, exploitation, reproduction, editing, distribution,<br>
as well as in the event of applications for industrial property rights.<br>
*****************************************************************************************************<br>
DESCRIPTION:<br>
Effective value of a SWITCH recipe field: TRUE for on (see m_Value).<br>
****************************************************************************************************)
METHOD m_Switch : BOOL
VAR_INPUT
	vi_un_Field							: UINT;	// [-] 1..the field count
END_VAR
m_Switch := m_Value(vi_un_Field := vi_un_Field) <> 0;
END_METHOD

(****************************************************************************************************<br>
© Syntegon Group.<br>
All rights reserved, also regarding any disposal, exploitation, reproduction, editing, distribution,<br>
as well as in the event of applications for industrial property rights.<br>
*****************************************************************************************************<br>
DESCRIPTION:<br>
Effective value of recipe field vi_un_Field, for the application's logic: the active recipe's, else the program<br>
value. 0 for a field not declared. A SWITCH gives 1 or 0, an INTEGER or CHOICE a whole number (m_Switch,<br>
m_Integer give them typed).<br>
****************************************************************************************************)
METHOD m_Value : LREAL
VAR_INPUT
	vi_un_Field							: UINT;	// [-] 1..the field count
END_VAR
IF vi_un_Field > 0 AND vi_un_Field <= vo_Config.nFieldCount THEN
	m_Value := vo_Config.aActive[vi_un_Field - 1];
ELSE
	m_Value := 0;
END_IF
END_METHOD

END_FUNCTION_BLOCK

// ---- POUs/_FB_ConfigComponent.TcPOU
(****************************************************************************************************<br>
© Syntegon Group.<br>
All rights reserved, also regarding any disposal, exploitation, reproduction, editing, distribution,<br>
as well as in the event of applications for industrial property rights.<br>
*****************************************************************************************************<br>
DESCRIPTION:<br>
Base of every parameter FB (_FB_ConfigConveyor, _FB_ConfigDelta, _FB_ConfigXtsGantry, ...): the config<br>
manifest entry, what is done with a staging (ADR 0017) and the helpers for zones, fingers, limit areas and<br>
track modules the derived FBs share. Not used directly.<br>
*****************************************************************************************************<br>
VERSION         ¦ DATE       ¦ NAME      ¦ CHANGE<br>
Syn_Config 1.0.0 ¦ 2026-11-10 ¦ J.Willner ¦ First version: conveyor and Delta<br>
Syn_Config 1.1.0 ¦ 2026-11-10 ¦ J.Willner ¦ Helpers m_PassOn..., m_Invalid... for every type<br>
Syn_Config 2.0.0 ¦ 2026-11-11 ¦ J.Willner ¦ m_InvalidFingers, m_PassOnFingers (ADR 0018)<br>
Syn_Config 2.3.0 ¦ 2026-11-14 ¦ J.Willner ¦ m_HandleStaging; symbol path from _FC_VisuSymbolPath<br>
Syn_Config 2.4.0 ¦ 2026-11-19 ¦ J.Willner ¦ m_Register: several id 0 entries told apart by path (topology FB)<br>
****************************************************************************************************)
{attribute 'reflection'}
FUNCTION_BLOCK ABSTRACT _FB_ConfigComponent
VAR
	udn_ComponentId						: UDINT;	// [-] id of the Syn_Visu component, 0 = not registered
	(* Device tree path of this instance, e.g. 'RPP_Visu.Syn_Visu_Demo.P_VisuDemoDelta.fb_InfeedParam', set by TwinCAT
	   at initialisation. *)
	{attribute 'instance-path'}
	{attribute 'noinit'}
	str_InstancePath					: STRING(255);
	str_SymbolPath						: STRING(255);	// symbol path of vo_Config for the manifest, from str_InstancePath
END_VAR

(****************************************************************************************************<br>
© Syntegon Group.<br>
All rights reserved, also regarding any disposal, exploitation, reproduction, editing, distribution,<br>
as well as in the event of applications for industrial property rights.<br>
*****************************************************************************************************<br>
DESCRIPTION:<br>
Type of the Syn_Visu component this FB parametrises. Overridden by every derived FB.<br>
****************************************************************************************************)
METHOD PROTECTED m_ComponentType : SynVisu.E_VisuComponentType
m_ComponentType := SynVisu.E_VisuComponentType.NONE;
END_METHOD

(****************************************************************************************************<br>
© Syntegon Group.<br>
All rights reserved, also regarding any disposal, exploitation, reproduction, editing, distribution,<br>
as well as in the event of applications for industrial property rights.<br>
*****************************************************************************************************<br>
DESCRIPTION:<br>
Reports the staging as handled: taken over (or reset) with an empty vi_str_Rejection, else rejected for that<br>
reason. Clears bStaged and bReset. TRUE when taken over.<br>
****************************************************************************************************)
METHOD PRIVATE m_Handled : BOOL
VAR_IN_OUT
	vio_Staging							: ST_ConfigStaging;	// vo_Config.stStaging
	vio_Status							: ST_ConfigStatus;	// vo_Config.stStatus
END_VAR
VAR_INPUT
	vi_str_Rejection					: STRING(80);	// why the set is not taken over; '' = taken over
END_VAR
m_Handled := vi_str_Rejection = '';
vio_Status.nHandledStageId := vio_Staging.nStageId;
IF m_Handled THEN
	vio_Status.eResult := E_ConfigResult.APPLIED;
	vio_Status.sMessage := '';
ELSE
	vio_Status.eResult := E_ConfigResult.REJECTED;
	vio_Status.sMessage := vi_str_Rejection;
END_IF
vio_Staging.bStaged := FALSE;
vio_Staging.bReset := FALSE;
END_METHOD

(****************************************************************************************************<br>
© Syntegon Group.<br>
All rights reserved, also regarding any disposal, exploitation, reproduction, editing, distribution,<br>
as well as in the event of applications for industrial property rights.<br>
*****************************************************************************************************<br>
DESCRIPTION:<br>
The staging lifecycle of every parameter FB (ADR 0017), for m_Cycle of the derived FB: a reset makes the active<br>
set invalid at once; a staged set waits while the application does not allow a take-over (PENDING), is rejected<br>
when based on another version than the active one or when m_InvalidStaged names a reason, and is taken over<br>
otherwise under a new version that never repeats. Reports the result in vio_Status, also the active version.<br>
The derived FB copies the staged set into its active set when vo_b_TakeOver says so.<br>
*****************************************************************************************************<br>
OUTPUT VALUES:<br>
TRUE in the cycle a set was taken over or reset.<br>
****************************************************************************************************)
METHOD PROTECTED m_HandleStaging : BOOL
VAR_IN_OUT
	vio_Staging							: ST_ConfigStaging;	// vo_Config.stStaging
	vio_Status							: ST_ConfigStatus;	// vo_Config.stStatus
	vio_b_Valid							: BOOL;	// the active set's bValid
	vio_udn_Version						: UDINT;	// [-] the active set's nVersion
	vio_udn_LastVersion					: UDINT;	// [-] the active set's nLastVersion
END_VAR
VAR_INPUT
	vi_b_ApplyAllowed					: BOOL;	// [-] the application allows taking a set over now
END_VAR
VAR_OUTPUT
	vo_b_TakeOver						: BOOL;	// TRUE: copy the staged set into the active set now
END_VAR
VAR
	udn_TempActiveVersion				: UDINT;	// [-] version of the active set, 0 = program values
	str_TempRejection					: STRING(80);
END_VAR
m_HandleStaging := FALSE;
vo_b_TakeOver := FALSE;
udn_TempActiveVersion := SEL(vio_b_Valid, 0, vio_udn_Version);
IF vio_Staging.bReset THEN
	vio_b_Valid := FALSE;
	m_Handled(vio_Staging := vio_Staging, vio_Status := vio_Status, vi_str_Rejection := '');
	m_HandleStaging := TRUE;
ELSIF vio_Staging.bStaged THEN
	IF NOT vi_b_ApplyAllowed THEN
		vio_Status.eResult := E_ConfigResult.PENDING;
	ELSIF vio_Staging.nBaseVersion <> udn_TempActiveVersion THEN
		m_Handled(vio_Staging := vio_Staging, vio_Status := vio_Status,
			vi_str_Rejection := CONCAT(CONCAT('Based on version ', UDINT_TO_STRING(vio_Staging.nBaseVersion)),
				CONCAT(', but version ', CONCAT(UDINT_TO_STRING(udn_TempActiveVersion), ' is active'))));
	ELSE
		str_TempRejection := m_InvalidStaged();
		IF str_TempRejection = '' THEN
			vio_udn_LastVersion := vio_udn_LastVersion + 1;
			vio_udn_Version := vio_udn_LastVersion;
			vio_b_Valid := TRUE;
			vo_b_TakeOver := TRUE;
			m_HandleStaging := TRUE;
		END_IF
		m_Handled(vio_Staging := vio_Staging, vio_Status := vio_Status, vi_str_Rejection := str_TempRejection);
	END_IF
END_IF
vio_Status.nActiveVersion := SEL(vio_b_Valid, 0, vio_udn_Version);
END_METHOD

(****************************************************************************************************<br>
© Syntegon Group.<br>
All rights reserved, also regarding any disposal, exploitation, reproduction, editing, distribution,<br>
as well as in the event of applications for industrial property rights.<br>
*****************************************************************************************************<br>
DESCRIPTION:<br>
Id given to m_Register (the Syn_Visu component's id); 0 while not registered.<br>
****************************************************************************************************)
METHOD m_Id : UDINT
m_Id := udn_ComponentId;
END_METHOD

(****************************************************************************************************<br>
© Syntegon Group.<br>
All rights reserved, also regarding any disposal, exploitation, reproduction, editing, distribution,<br>
as well as in the event of applications for industrial property rights.<br>
*****************************************************************************************************<br>
DESCRIPTION:<br>
Why a staged set's gripper fingers cannot be taken over; '' when they can: more fingers than the list holds, or<br>
a finger without a diameter or height.<br>
****************************************************************************************************)
METHOD PROTECTED m_InvalidFingers : STRING(80)
VAR_IN_OUT CONSTANT
	(* staged fingers *)
	vio_aFingers						: ARRAY[0..SynVisu.VISU_GlobalConst_Param.VISU_un_MAX_FINGERS - 1] OF SynVisu.ST_VisuFinger;
END_VAR
VAR_INPUT
	vi_un_Count							: UINT;	// [-] staged fingers in vio_aFingers
END_VAR
VAR
	un_TempIndex						: UINT;
END_VAR
m_InvalidFingers := '';
IF vi_un_Count > SynVisu.VISU_GlobalConst_Param.VISU_un_MAX_FINGERS THEN
	m_InvalidFingers := CONCAT('More than ', CONCAT(UINT_TO_STRING(SynVisu.VISU_GlobalConst_Param.VISU_un_MAX_FINGERS), ' fingers'));
	RETURN;
END_IF
un_TempIndex := 0;
WHILE un_TempIndex < vi_un_Count DO
	IF vio_aFingers[un_TempIndex].fDiameter <= 0 OR vio_aFingers[un_TempIndex].fHeight <= 0 THEN
		m_InvalidFingers := CONCAT('Finger ', CONCAT(UINT_TO_STRING(un_TempIndex + 1), ' has no diameter or height'));
		RETURN;
	END_IF
	un_TempIndex := un_TempIndex + 1;
END_WHILE
END_METHOD

(****************************************************************************************************<br>
© Syntegon Group.<br>
All rights reserved, also regarding any disposal, exploitation, reproduction, editing, distribution,<br>
as well as in the event of applications for industrial property rights.<br>
*****************************************************************************************************<br>
DESCRIPTION:<br>
Why a staged set's track modules cannot be taken over; '' when they can: more modules than the list holds,<br>
none at all, or a module without a length.<br>
****************************************************************************************************)
METHOD PROTECTED m_InvalidModules : STRING(80)
VAR_IN_OUT CONSTANT
	(* staged modules *)
	vio_aModules						: ARRAY[0..SynVisu.VISU_GlobalConst_Param.VISU_un_MAX_MODULES - 1] OF SynVisu.ST_VisuTrackModule;
END_VAR
VAR_INPUT
	vi_un_Count							: UINT;	// [-] staged modules in vio_aModules
END_VAR
VAR
	un_TempIndex						: UINT;
END_VAR
m_InvalidModules := '';
IF vi_un_Count > SynVisu.VISU_GlobalConst_Param.VISU_un_MAX_MODULES THEN
	m_InvalidModules := CONCAT('More than ', CONCAT(UINT_TO_STRING(SynVisu.VISU_GlobalConst_Param.VISU_un_MAX_MODULES), ' track modules'));
	RETURN;
END_IF
IF vi_un_Count = 0 THEN
	m_InvalidModules := 'A track without modules';
	RETURN;
END_IF
un_TempIndex := 0;
WHILE un_TempIndex < vi_un_Count DO
	IF vio_aModules[un_TempIndex].fLength <= 0 THEN
		m_InvalidModules := CONCAT('Track module ', CONCAT(UINT_TO_STRING(un_TempIndex + 1), ' has no length'));
		RETURN;
	END_IF
	un_TempIndex := un_TempIndex + 1;
END_WHILE
END_METHOD

(****************************************************************************************************<br>
© Syntegon Group.<br>
All rights reserved, also regarding any disposal, exploitation, reproduction, editing, distribution,<br>
as well as in the event of applications for industrial property rights.<br>
*****************************************************************************************************<br>
DESCRIPTION:<br>
Why the set in vo_Config.stStaged cannot be taken over; '' when it can. Each parameter FB names its own checks;<br>
m_HandleStaging asks before a take-over.<br>
****************************************************************************************************)
METHOD PROTECTED ABSTRACT m_InvalidStaged : STRING(80)
END_METHOD

(****************************************************************************************************<br>
© Syntegon Group.<br>
All rights reserved, also regarding any disposal, exploitation, reproduction, editing, distribution,<br>
as well as in the event of applications for industrial property rights.<br>
*****************************************************************************************************<br>
DESCRIPTION:<br>
Why a staged set's zones cannot be taken over; '' when they can: more zones than the list holds, or a zone on<br>
no conveyor (id 0).<br>
****************************************************************************************************)
METHOD PROTECTED m_InvalidZones : STRING(80)
VAR_IN_OUT CONSTANT
	(* staged zones *)
	vio_aZones							: ARRAY[0..SynVisu.VISU_GlobalConst_Param.VISU_un_MAX_ZONES - 1] OF SynVisu.ST_VisuZone;
END_VAR
VAR_INPUT
	vi_un_Count							: UINT;	// [-] staged zones in vio_aZones
END_VAR
VAR
	un_TempIndex						: UINT;
END_VAR
m_InvalidZones := '';
IF vi_un_Count > SynVisu.VISU_GlobalConst_Param.VISU_un_MAX_ZONES THEN
	m_InvalidZones := CONCAT('More than ', CONCAT(UINT_TO_STRING(SynVisu.VISU_GlobalConst_Param.VISU_un_MAX_ZONES), ' zones'));
	RETURN;
END_IF
un_TempIndex := 0;
WHILE un_TempIndex < vi_un_Count DO
	IF vio_aZones[un_TempIndex].nConveyorId = 0 THEN
		m_InvalidZones := CONCAT('Zone ', CONCAT(UINT_TO_STRING(un_TempIndex + 1), ' lies on no conveyor'));
		RETURN;
	END_IF
	un_TempIndex := un_TempIndex + 1;
END_WHILE
END_METHOD

(****************************************************************************************************<br>
© Syntegon Group.<br>
All rights reserved, also regarding any disposal, exploitation, reproduction, editing, distribution,<br>
as well as in the event of applications for industrial property rights.<br>
*****************************************************************************************************<br>
DESCRIPTION:<br>
Passes the effective gripper fingers with their flange offsets on to a robot's Syn_Visu FB (ADR 0018). Syn_Visu's<br>
finger count only grows: the fingers are cleared first only when the set has fewer than the visualisation, so<br>
its config version only changes when a value does.<br>
****************************************************************************************************)
METHOD PROTECTED m_PassOnFingers : BOOL
VAR_IN_OUT
	vio_Visu							: SynVisu._FB_VisuRobot;	// the robot's Syn_Visu FB
END_VAR
VAR_IN_OUT CONSTANT
	(* effective fingers *)
	vio_aFingers						: ARRAY[0..SynVisu.VISU_GlobalConst_Param.VISU_un_MAX_FINGERS - 1] OF SynVisu.ST_VisuFinger;
END_VAR
VAR_INPUT
	vi_un_Count							: UINT;	// [-] effective fingers in vio_aFingers
	vi_un_VisuCount						: UINT;	// [-] fingers the visualisation has now, its stConfig.nFingerCount
END_VAR
VAR
	un_TempIndex						: UINT;
END_VAR
m_PassOnFingers := TRUE;
IF vi_un_VisuCount > vi_un_Count THEN
	vio_Visu.m_ClearFingers();
END_IF
un_TempIndex := 0;
WHILE un_TempIndex < vi_un_Count AND un_TempIndex < SynVisu.VISU_GlobalConst_Param.VISU_un_MAX_FINGERS DO
	vio_Visu.m_SetFinger(vi_un_Finger := un_TempIndex + 1, vi_lr_Diameter := vio_aFingers[un_TempIndex].fDiameter,
		vi_lr_Height := vio_aFingers[un_TempIndex].fHeight);
	vio_Visu.m_SetFingerOffset(vi_un_Finger := un_TempIndex + 1, vi_lr_X := vio_aFingers[un_TempIndex].stOffset.fX,
		vi_lr_Y := vio_aFingers[un_TempIndex].stOffset.fY, vi_lr_Z := vio_aFingers[un_TempIndex].stOffset.fZ,
		vi_lr_Rz := vio_aFingers[un_TempIndex].stOffset.fRz);
	un_TempIndex := un_TempIndex + 1;
END_WHILE
END_METHOD

(****************************************************************************************************<br>
© Syntegon Group.<br>
All rights reserved, also regarding any disposal, exploitation, reproduction, editing, distribution,<br>
as well as in the event of applications for industrial property rights.<br>
*****************************************************************************************************<br>
DESCRIPTION:<br>
Passes the effective limit area and TCP limit area on to a robot's Syn_Visu FB (Delta, XTS gantry, Cartesian);<br>
an area with bActive = FALSE is cleared.<br>
****************************************************************************************************)
METHOD PROTECTED m_PassOnLimitAreas : BOOL
VAR_IN_OUT
	vio_Visu							: SynVisu._FB_VisuRobot;	// the robot's Syn_Visu FB
END_VAR
VAR_IN_OUT CONSTANT
	vio_LimitArea						: SynVisu.ST_VisuLimitArea;	// effective limit area
	vio_TcpLimitArea					: SynVisu.ST_VisuLimitArea;	// effective TCP limit area
END_VAR
m_PassOnLimitAreas := TRUE;
IF vio_LimitArea.bActive THEN
	vio_Visu.m_SetLimitArea(vi_lr_XMin := vio_LimitArea.fXMin, vi_lr_XMax := vio_LimitArea.fXMax,
		vi_lr_YMin := vio_LimitArea.fYMin, vi_lr_YMax := vio_LimitArea.fYMax,
		vi_lr_ZMin := vio_LimitArea.fZMin, vi_lr_ZMax := vio_LimitArea.fZMax);
ELSE
	vio_Visu.m_ClearLimitArea();
END_IF
IF vio_TcpLimitArea.bActive THEN
	vio_Visu.m_SetTcpLimitArea(vi_lr_XMin := vio_TcpLimitArea.fXMin, vi_lr_XMax := vio_TcpLimitArea.fXMax,
		vi_lr_YMin := vio_TcpLimitArea.fYMin, vi_lr_YMax := vio_TcpLimitArea.fYMax,
		vi_lr_ZMin := vio_TcpLimitArea.fZMin, vi_lr_ZMax := vio_TcpLimitArea.fZMax);
ELSE
	vio_Visu.m_ClearTcpLimitArea();
END_IF
END_METHOD

(****************************************************************************************************<br>
© Syntegon Group.<br>
All rights reserved, also regarding any disposal, exploitation, reproduction, editing, distribution,<br>
as well as in the event of applications for industrial property rights.<br>
*****************************************************************************************************<br>
DESCRIPTION:<br>
Passes the effective track modules on to an XTS track's Syn_Visu FB (XTS gantry, XTS loop). Syn_Visu's module<br>
count only grows: the modules are cleared first only when the set has fewer than the visualisation, so its<br>
config version only changes when a value does.<br>
****************************************************************************************************)
METHOD PROTECTED m_PassOnModules : BOOL
VAR_IN_OUT
	vio_Visu							: SynVisu._FB_VisuXtsTrack;	// the track's Syn_Visu FB
END_VAR
VAR_IN_OUT CONSTANT
	(* effective modules *)
	vio_aModules						: ARRAY[0..SynVisu.VISU_GlobalConst_Param.VISU_un_MAX_MODULES - 1] OF SynVisu.ST_VisuTrackModule;
END_VAR
VAR_INPUT
	vi_un_Count							: UINT;	// [-] effective modules in vio_aModules
	vi_un_VisuCount						: UINT;	// [-] modules the visualisation has now, its stConfig.nModuleCount
END_VAR
VAR
	un_TempIndex						: UINT;
END_VAR
m_PassOnModules := TRUE;
IF vi_un_VisuCount > vi_un_Count THEN
	vio_Visu.m_ClearModules();
END_IF
un_TempIndex := 0;
WHILE un_TempIndex < vi_un_Count AND un_TempIndex < SynVisu.VISU_GlobalConst_Param.VISU_un_MAX_MODULES DO
	vio_Visu.m_SetModule(vi_un_Module := un_TempIndex + 1, vi_e_Kind := vio_aModules[un_TempIndex].eKind,
		vi_lr_Length := vio_aModules[un_TempIndex].fLength);
	un_TempIndex := un_TempIndex + 1;
END_WHILE
END_METHOD

(****************************************************************************************************<br>
© Syntegon Group.<br>
All rights reserved, also regarding any disposal, exploitation, reproduction, editing, distribution,<br>
as well as in the event of applications for industrial property rights.<br>
*****************************************************************************************************<br>
DESCRIPTION:<br>
Passes the effective zones on to a Syn_Visu component with zones (robot, detector, station). Syn_Visu's zone<br>
count only grows: the zones are cleared first only when the set has fewer than the visualisation, so its<br>
config version only changes when a value does.<br>
****************************************************************************************************)
METHOD PROTECTED m_PassOnZones : BOOL
VAR_IN_OUT
	vio_Visu							: SynVisu._FB_VisuZoneComponent;	// the component's Syn_Visu FB
END_VAR
VAR_IN_OUT CONSTANT
	(* effective zones *)
	vio_aZones							: ARRAY[0..SynVisu.VISU_GlobalConst_Param.VISU_un_MAX_ZONES - 1] OF SynVisu.ST_VisuZone;
END_VAR
VAR_INPUT
	vi_un_Count							: UINT;	// [-] effective zones in vio_aZones
	vi_un_VisuCount						: UINT;	// [-] zones the visualisation has now, its stConfig.nZoneCount
END_VAR
VAR
	un_TempIndex						: UINT;
END_VAR
m_PassOnZones := TRUE;
IF vi_un_VisuCount > vi_un_Count THEN
	vio_Visu.m_ClearZones();
END_IF
un_TempIndex := 0;
WHILE un_TempIndex < vi_un_Count AND un_TempIndex < SynVisu.VISU_GlobalConst_Param.VISU_un_MAX_ZONES DO
	vio_Visu.m_SetZone(vi_un_Zone := un_TempIndex + 1, vi_udn_ConveyorId := vio_aZones[un_TempIndex].nConveyorId,
		vi_lr_Start := vio_aZones[un_TempIndex].fStart, vi_lr_End := vio_aZones[un_TempIndex].fEnd,
		vi_lr_AllocationOffset := vio_aZones[un_TempIndex].fAllocationOffset,
		vi_lr_CcsOffset := vio_aZones[un_TempIndex].fCcsOffset,
		vi_lr_StartY := vio_aZones[un_TempIndex].fStartY, vi_lr_EndY := vio_aZones[un_TempIndex].fEndY);
	un_TempIndex := un_TempIndex + 1;
END_WHILE
END_METHOD

(****************************************************************************************************<br>
© Syntegon Group.<br>
All rights reserved, also regarding any disposal, exploitation, reproduction, editing, distribution,<br>
as well as in the event of applications for industrial property rights.<br>
*****************************************************************************************************<br>
DESCRIPTION:<br>
Adds this parameter FB to the config manifest under the id of the Syn_Visu component it parametrises.<br>
Idempotent: call it every cycle. The symbol path the gateway reads comes from the instance's own path, as in<br>
Syn_Visu (VISU_un_INSTANCE_PATH_SKIP).<br>
*****************************************************************************************************<br>
OUTPUT VALUES:<br>
FALSE for vi_udn_Id = 0 (but for _FB_ConfigMachine and _FB_ConfigTopology, which register with id 0 and are told<br>
apart by their path), an id already used by a different entry, or a full manifest.<br>
****************************************************************************************************)
METHOD m_Register : BOOL
VAR_IN_OUT
	vio_Manifest						: ST_ConfigManifest;	// GVL_Config.stManifest of the application
END_VAR
VAR_INPUT
	vi_udn_Id							: UDINT;	// [-] id of the Syn_Visu component, e.g. fb_Infeed.m_Id()
END_VAR
VAR
	e_TempType							: SynVisu.E_VisuComponentType;
	un_TempIndex						: UINT;
END_VAR
m_Register := FALSE;
(* Always report the contract version of the library actually running, also after an online change. *)
vio_Manifest.nProtocolVersion := CONFIG_GlobalConst.CONFIG_un_PROTOCOL_VERSION;
vio_Manifest.sLibraryVersion := CONFIG_GlobalConst.CONFIG_str_LIBRARY_VERSION;
e_TempType := m_ComponentType();
(* Id 0 is the machine-wide FBs', whose type is NONE (_FB_ConfigMachine, _FB_ConfigTopology); every parameter FB has a
   component's id. *)
IF (vi_udn_Id = 0) <> (e_TempType = SynVisu.E_VisuComponentType.NONE) THEN
	RETURN;
END_IF
IF str_SymbolPath = '' THEN
	str_SymbolPath := SynVisu._FC_VisuSymbolPath(vio_str_InstancePath := str_InstancePath, vi_str_Member := '.vo_Config');
END_IF

(* An existing entry with the same id must match exactly. Id 0 is shared by the machine-wide FBs (machine and
   topology), told apart by their path. *)
un_TempIndex := 0;
WHILE un_TempIndex < vio_Manifest.nCount AND un_TempIndex < CONFIG_GlobalConst_Param.CONFIG_un_MAX_MANIFEST_ENTRIES DO
	IF vio_Manifest.aEntries[un_TempIndex].nId = vi_udn_Id
		AND (vi_udn_Id <> 0 OR vio_Manifest.aEntries[un_TempIndex].sPath = str_SymbolPath)
	THEN
		m_Register := vio_Manifest.aEntries[un_TempIndex].eType = e_TempType
					AND vio_Manifest.aEntries[un_TempIndex].sPath = str_SymbolPath;
		IF m_Register THEN
			udn_ComponentId := vi_udn_Id;
		END_IF
		RETURN;
	END_IF
	un_TempIndex := un_TempIndex + 1;
END_WHILE

(* New entry. *)
IF vio_Manifest.nCount >= CONFIG_GlobalConst_Param.CONFIG_un_MAX_MANIFEST_ENTRIES THEN
	RETURN;
END_IF
vio_Manifest.aEntries[vio_Manifest.nCount].nId := vi_udn_Id;
vio_Manifest.aEntries[vio_Manifest.nCount].eType := e_TempType;
vio_Manifest.aEntries[vio_Manifest.nCount].sPath := str_SymbolPath;
vio_Manifest.nCount := vio_Manifest.nCount + 1;
udn_ComponentId := vi_udn_Id;
m_Register := TRUE;
END_METHOD

END_FUNCTION_BLOCK

// ---- POUs/_FB_ConfigTopology.TcPOU
(****************************************************************************************************<br>
© Syntegon Group.<br>
All rights reserved, also regarding any disposal, exploitation, reproduction, editing, distribution,<br>
as well as in the event of applications for industrial property rights.<br>
*****************************************************************************************************<br>
DESCRIPTION:<br>
The machine's topology (config protocol 5, ADR 0023): how the parts of the application relate. The application<br>
declares the kinds of its topology nodes, the roles a link may have, every node of its full build-out with the<br>
Syn_Visu components it stands for, and its root node; its program values are the parents and links it uses. One per<br>
application, listed in the config manifest with id 0 like the machine FB. Typical cycle:<br>
  fb_Topology.m_Register(vio_Manifest := GVL_Config.stManifest, vi_udn_Id := 0);<br>
  fb_Topology.m_DeclareKind(vi_un_Kind := 1, vi_str_Name := 'Line');<br>
  fb_Topology.m_DeclareKind(vi_un_Kind := 2, vi_str_Name := 'PPH');<br>
  fb_Topology.m_AllowParent(vi_un_Kind := 2, vi_un_ParentKind := 1);<br>
  fb_Topology.m_DeclareRole(vi_un_Role := 1, vi_str_Name := 'Infeed1', vi_un_HolderKind := 2, vi_b_Required := TRUE);<br>
  fb_Topology.m_AllowTarget(vi_un_Role := 1, vi_un_TargetKind := 3);<br>
  fb_Topology.m_DeclareNode(vi_dn_Id := 21, vi_str_Name := 'PPH1', vi_un_Kind := 2);<br>
  fb_Topology.m_AddComponent(vi_dn_Node := 21, vi_udn_ComponentId := fb_Delta1.m_Id());<br>
  fb_Topology.m_SetRoot(vi_dn_Node := 1);<br>
  fb_Topology.m_SetParent(vi_dn_Node := 21, vi_dn_Parent := 1);<br>
  fb_Topology.m_Link(vi_dn_Node := 21, vi_un_Role := 1, vi_dn_Target := 30);<br>
  fb_Topology.m_Cycle();<br>
*****************************************************************************************************<br>
OUTPUT VALUES:<br>
vo_Config is the contract structure the gateway reads at the path in the config manifest.<br>
*****************************************************************************************************<br>
LIMITS:<br>
CONFIG_un_MAX_TOPOLOGY_KINDS kinds, CONFIG_un_MAX_TOPOLOGY_ROLES roles, CONFIG_un_MAX_TOPOLOGY_NODES nodes,<br>
CONFIG_un_MAX_TOPOLOGY_LINKS links, CONFIG_un_MAX_NODE_COMPONENTS components per node. The gateway reads the<br>
declaration when it discovers the PLC: declare everything from the start.<br>
*****************************************************************************************************<br>
VERSION         ¦ DATE       ¦ NAME      ¦ CHANGE<br>
Syn_Config 2.4.0 ¦ 2026-11-19 ¦ J.Willner ¦ Created: declaration and program values (protocol 5, #56)<br>
****************************************************************************************************)
FUNCTION_BLOCK _FB_ConfigTopology EXTENDS _FB_ConfigComponent
VAR_OUTPUT
	vo_Config							: ST_ConfigTopology;	// contract structure of the gateway
END_VAR
VAR
	ProgramLinks						: ST_ConfigTopologyLinks;	// the program values, given with m_SetParent and m_Link
END_VAR

(****************************************************************************************************<br>
© Syntegon Group.<br>
All rights reserved, also regarding any disposal, exploitation, reproduction, editing, distribution,<br>
as well as in the event of applications for industrial property rights.<br>
*****************************************************************************************************<br>
DESCRIPTION:<br>
Names a Syn_Visu component the declared node vi_dn_Node stands for, e.g. a PPH's Delta robot. Idempotent: call it<br>
every cycle with m_DeclareNode.<br>
*****************************************************************************************************<br>
OUTPUT VALUES:<br>
FALSE for a node not declared, component id 0, or more than CONFIG_un_MAX_NODE_COMPONENTS components.<br>
****************************************************************************************************)
METHOD m_AddComponent : BOOL
VAR_INPUT
	vi_dn_Node							: DINT;	// [-] the node's id
	vi_udn_ComponentId					: UDINT;	// [-] manifest id of the Syn_Visu component, e.g. fb_Delta1.m_Id()
END_VAR
VAR
	n_TempNode							: INT;
	un_TempIndex						: UINT;
END_VAR
n_TempNode := m_NodeIndex(vi_dn_Id := vi_dn_Node);
m_AddComponent := n_TempNode >= 0 AND vi_udn_ComponentId <> 0;
IF NOT m_AddComponent THEN
	RETURN;
END_IF
un_TempIndex := 0;
WHILE un_TempIndex < vo_Config.aNodes[n_TempNode].nComponentCount
	AND un_TempIndex < CONFIG_GlobalConst_Param.CONFIG_un_MAX_NODE_COMPONENTS
DO
	IF vo_Config.aNodes[n_TempNode].aComponents[un_TempIndex] = vi_udn_ComponentId THEN
		RETURN;
	END_IF
	un_TempIndex := un_TempIndex + 1;
END_WHILE
IF vo_Config.aNodes[n_TempNode].nComponentCount >= CONFIG_GlobalConst_Param.CONFIG_un_MAX_NODE_COMPONENTS THEN
	m_AddComponent := FALSE;
	RETURN;
END_IF
vo_Config.aNodes[n_TempNode].aComponents[vo_Config.aNodes[n_TempNode].nComponentCount] := vi_udn_ComponentId;
vo_Config.aNodes[n_TempNode].nComponentCount := vo_Config.aNodes[n_TempNode].nComponentCount + 1;
END_METHOD

(****************************************************************************************************<br>
© Syntegon Group.<br>
All rights reserved, also regarding any disposal, exploitation, reproduction, editing, distribution,<br>
as well as in the event of applications for industrial property rights.<br>
*****************************************************************************************************<br>
DESCRIPTION:<br>
Allows a node of kind vi_un_ParentKind to be the parent of a node of kind vi_un_Kind, e.g. a cell the parent of a<br>
PPH. Idempotent: call it every cycle with m_DeclareKind.<br>
*****************************************************************************************************<br>
OUTPUT VALUES:<br>
FALSE when either kind is not declared.<br>
****************************************************************************************************)
METHOD m_AllowParent : BOOL
VAR_INPUT
	vi_un_Kind							: UINT;	// [-] the child's kind, 1..its count
	vi_un_ParentKind					: UINT;	// [-] the parent's kind, 1..its count
END_VAR
m_AllowParent := vi_un_Kind > 0 AND vi_un_Kind <= vo_Config.nKindCount
	AND vi_un_ParentKind > 0 AND vi_un_ParentKind <= vo_Config.nKindCount;
IF NOT m_AllowParent THEN
	RETURN;
END_IF
vo_Config.aKinds[vi_un_Kind - 1].nParentKinds := vo_Config.aKinds[vi_un_Kind - 1].nParentKinds
	OR SHL(DWORD#1, vi_un_ParentKind - 1);
END_METHOD

(****************************************************************************************************<br>
© Syntegon Group.<br>
All rights reserved, also regarding any disposal, exploitation, reproduction, editing, distribution,<br>
as well as in the event of applications for industrial property rights.<br>
*****************************************************************************************************<br>
DESCRIPTION:<br>
Allows a link in role vi_un_Role to point to a node of kind vi_un_TargetKind, e.g. Infeed1 to a transport.<br>
Idempotent: call it every cycle with m_DeclareRole.<br>
*****************************************************************************************************<br>
OUTPUT VALUES:<br>
FALSE when the role or the kind is not declared.<br>
****************************************************************************************************)
METHOD m_AllowTarget : BOOL
VAR_INPUT
	vi_un_Role							: UINT;	// [-] the role, 1..its count
	vi_un_TargetKind					: UINT;	// [-] the kind it may point to, 1..its count
END_VAR
m_AllowTarget := vi_un_Role > 0 AND vi_un_Role <= vo_Config.nRoleCount
	AND vi_un_TargetKind > 0 AND vi_un_TargetKind <= vo_Config.nKindCount;
IF NOT m_AllowTarget THEN
	RETURN;
END_IF
vo_Config.aRoles[vi_un_Role - 1].nTargetKinds := vo_Config.aRoles[vi_un_Role - 1].nTargetKinds
	OR SHL(DWORD#1, vi_un_TargetKind - 1);
END_METHOD

(****************************************************************************************************<br>
© Syntegon Group.<br>
All rights reserved, also regarding any disposal, exploitation, reproduction, editing, distribution,<br>
as well as in the event of applications for industrial property rights.<br>
*****************************************************************************************************<br>
DESCRIPTION:<br>
Every cycle, after the declaration and the program values: gives the links in effect in vo_Config.stActive, the<br>
program values.<br>
*****************************************************************************************************<br>
OUTPUT VALUES:<br>
TRUE.<br>
****************************************************************************************************)
METHOD m_Cycle : BOOL
vo_Config.stActive := ProgramLinks;
m_Cycle := TRUE;
END_METHOD

(****************************************************************************************************<br>
© Syntegon Group.<br>
All rights reserved, also regarding any disposal, exploitation, reproduction, editing, distribution,<br>
as well as in the event of applications for industrial property rights.<br>
*****************************************************************************************************<br>
DESCRIPTION:<br>
Declares kind vi_un_Kind (1..CONFIG_un_MAX_TOPOLOGY_KINDS) of topology node, e.g. 'PPH' or 'Transport'. Kinds are<br>
listed up to the highest one declared. Idempotent: call it every cycle, before the roles and nodes.<br>
*****************************************************************************************************<br>
OUTPUT VALUES:<br>
FALSE for vi_un_Kind = 0 or above CONFIG_un_MAX_TOPOLOGY_KINDS.<br>
****************************************************************************************************)
METHOD m_DeclareKind : BOOL
VAR_INPUT
	vi_un_Kind							: UINT;	// [-] 1..CONFIG_un_MAX_TOPOLOGY_KINDS
	vi_str_Name							: STRING(31);	// unique in the topology, e.g. 'PPH'
END_VAR
m_DeclareKind := vi_un_Kind > 0 AND vi_un_Kind <= CONFIG_GlobalConst_Param.CONFIG_un_MAX_TOPOLOGY_KINDS;
IF NOT m_DeclareKind THEN
	RETURN;
END_IF
vo_Config.aKinds[vi_un_Kind - 1].sName := vi_str_Name;
IF vi_un_Kind > vo_Config.nKindCount THEN
	vo_Config.nKindCount := vi_un_Kind;
END_IF
END_METHOD

(****************************************************************************************************<br>
© Syntegon Group.<br>
All rights reserved, also regarding any disposal, exploitation, reproduction, editing, distribution,<br>
as well as in the event of applications for industrial property rights.<br>
*****************************************************************************************************<br>
DESCRIPTION:<br>
Declares the topology node vi_dn_Id of the full build-out, in use or not, with its name and kind; nodes are listed<br>
in the order they are first declared. Idempotent: call it every cycle, after m_DeclareKind.<br>
*****************************************************************************************************<br>
OUTPUT VALUES:<br>
FALSE for id 0, a kind not declared, or more than CONFIG_un_MAX_TOPOLOGY_NODES nodes.<br>
****************************************************************************************************)
METHOD m_DeclareNode : BOOL
VAR_INPUT
	vi_dn_Id							: DINT;	// [-] the application's id, e.g. its context id; not 0
	vi_str_Name							: STRING(31);	// e.g. 'PPH1'
	vi_un_Kind							: UINT;	// [-] its kind, 1..the kind count
END_VAR
VAR
	n_TempIndex							: INT;
END_VAR
m_DeclareNode := vi_dn_Id <> 0 AND vi_un_Kind > 0 AND vi_un_Kind <= vo_Config.nKindCount;
IF NOT m_DeclareNode THEN
	RETURN;
END_IF
n_TempIndex := m_NodeIndex(vi_dn_Id := vi_dn_Id);
IF n_TempIndex < 0 THEN
	IF vo_Config.nNodeCount >= CONFIG_GlobalConst_Param.CONFIG_un_MAX_TOPOLOGY_NODES THEN
		m_DeclareNode := FALSE;
		RETURN;
	END_IF
	n_TempIndex := UINT_TO_INT(vo_Config.nNodeCount);
	vo_Config.nNodeCount := vo_Config.nNodeCount + 1;
	vo_Config.aNodes[n_TempIndex].nId := vi_dn_Id;
END_IF
vo_Config.aNodes[n_TempIndex].sName := vi_str_Name;
vo_Config.aNodes[n_TempIndex].nKind := vi_un_Kind;
END_METHOD

(****************************************************************************************************<br>
© Syntegon Group.<br>
All rights reserved, also regarding any disposal, exploitation, reproduction, editing, distribution,<br>
as well as in the event of applications for industrial property rights.<br>
*****************************************************************************************************<br>
DESCRIPTION:<br>
Declares role vi_un_Role (1..CONFIG_un_MAX_TOPOLOGY_ROLES) a link may have, e.g. 'Infeed1' held by a PPH; the kinds<br>
it may point to are allowed with m_AllowTarget. Roles are listed up to the highest one declared. The parent is no<br>
role (m_SetParent). Idempotent: call it every cycle, after m_DeclareKind.<br>
*****************************************************************************************************<br>
OUTPUT VALUES:<br>
FALSE for vi_un_Role = 0 or above CONFIG_un_MAX_TOPOLOGY_ROLES, or a holder kind not declared.<br>
****************************************************************************************************)
METHOD m_DeclareRole : BOOL
VAR_INPUT
	vi_un_Role							: UINT;	// [-] 1..CONFIG_un_MAX_TOPOLOGY_ROLES
	vi_str_Name							: STRING(31);	// unique in the topology, e.g. 'Infeed1'
	vi_un_HolderKind					: UINT;	// [-] the kind of node that holds the role
	vi_b_Required						: BOOL;	// a node in use of that kind must have a link in this role
END_VAR
m_DeclareRole := vi_un_Role > 0 AND vi_un_Role <= CONFIG_GlobalConst_Param.CONFIG_un_MAX_TOPOLOGY_ROLES
	AND vi_un_HolderKind > 0 AND vi_un_HolderKind <= vo_Config.nKindCount;
IF NOT m_DeclareRole THEN
	RETURN;
END_IF
vo_Config.aRoles[vi_un_Role - 1].sName := vi_str_Name;
vo_Config.aRoles[vi_un_Role - 1].nHolderKind := vi_un_HolderKind;
vo_Config.aRoles[vi_un_Role - 1].bRequired := vi_b_Required;
IF vi_un_Role > vo_Config.nRoleCount THEN
	vo_Config.nRoleCount := vi_un_Role;
END_IF
END_METHOD

(****************************************************************************************************<br>
© Syntegon Group.<br>
All rights reserved, also regarding any disposal, exploitation, reproduction, editing, distribution,<br>
as well as in the event of applications for industrial property rights.<br>
*****************************************************************************************************<br>
DESCRIPTION:<br>
The topology is not staged yet (config protocol 5 has no topology staging): nothing to reject.<br>
****************************************************************************************************)
METHOD PROTECTED m_InvalidStaged : STRING(80)
m_InvalidStaged := '';
END_METHOD

(****************************************************************************************************<br>
© Syntegon Group.<br>
All rights reserved, also regarding any disposal, exploitation, reproduction, editing, distribution,<br>
as well as in the event of applications for industrial property rights.<br>
*****************************************************************************************************<br>
DESCRIPTION:<br>
A program value: node vi_dn_Node points to node vi_dn_Target in role vi_un_Role, e.g. PPH1's Infeed1 is TBL1. A<br>
node has one link per role; linking it again in that role replaces the target. Role 0 is the parent<br>
(m_SetParent). Idempotent: call it every cycle after the declaration, before m_Cycle.<br>
*****************************************************************************************************<br>
OUTPUT VALUES:<br>
FALSE for a node, target or role not declared, or more than CONFIG_un_MAX_TOPOLOGY_LINKS links.<br>
****************************************************************************************************)
METHOD m_Link : BOOL
VAR_INPUT
	vi_dn_Node							: DINT;	// [-] id of the node that holds the link
	vi_un_Role							: UINT;	// [-] its role, 1..the role count; 0 = the parent
	vi_dn_Target						: DINT;	// [-] id of the node it points to
END_VAR
VAR
	un_TempIndex						: UINT;
END_VAR
m_Link := m_NodeIndex(vi_dn_Id := vi_dn_Node) >= 0 AND m_NodeIndex(vi_dn_Id := vi_dn_Target) >= 0
	AND vi_un_Role <= vo_Config.nRoleCount;
IF NOT m_Link THEN
	RETURN;
END_IF

(* The node's link in this role, if it has one. *)
un_TempIndex := 0;
WHILE un_TempIndex < ProgramLinks.nLinkCount AND un_TempIndex < CONFIG_GlobalConst_Param.CONFIG_un_MAX_TOPOLOGY_LINKS DO
	IF ProgramLinks.aLinks[un_TempIndex].nNode = vi_dn_Node AND ProgramLinks.aLinks[un_TempIndex].nRole = vi_un_Role THEN
		ProgramLinks.aLinks[un_TempIndex].nTarget := vi_dn_Target;
		RETURN;
	END_IF
	un_TempIndex := un_TempIndex + 1;
END_WHILE

(* New link. *)
IF ProgramLinks.nLinkCount >= CONFIG_GlobalConst_Param.CONFIG_un_MAX_TOPOLOGY_LINKS THEN
	m_Link := FALSE;
	RETURN;
END_IF
ProgramLinks.aLinks[ProgramLinks.nLinkCount].nNode := vi_dn_Node;
ProgramLinks.aLinks[ProgramLinks.nLinkCount].nRole := vi_un_Role;
ProgramLinks.aLinks[ProgramLinks.nLinkCount].nTarget := vi_dn_Target;
ProgramLinks.nLinkCount := ProgramLinks.nLinkCount + 1;
END_METHOD

(****************************************************************************************************<br>
© Syntegon Group.<br>
All rights reserved, also regarding any disposal, exploitation, reproduction, editing, distribution,<br>
as well as in the event of applications for industrial property rights.<br>
*****************************************************************************************************<br>
DESCRIPTION:<br>
Index in vo_Config.aNodes of the node with id vi_dn_Id; -1 when none is declared.<br>
****************************************************************************************************)
METHOD PRIVATE m_NodeIndex : INT
VAR_INPUT
	vi_dn_Id							: DINT;	// [-] the node's id
END_VAR
VAR
	un_TempIndex						: UINT;
END_VAR
m_NodeIndex := -1;
un_TempIndex := 0;
WHILE un_TempIndex < vo_Config.nNodeCount AND un_TempIndex < CONFIG_GlobalConst_Param.CONFIG_un_MAX_TOPOLOGY_NODES DO
	IF vo_Config.aNodes[un_TempIndex].nId = vi_dn_Id THEN
		m_NodeIndex := UINT_TO_INT(un_TempIndex);
		RETURN;
	END_IF
	un_TempIndex := un_TempIndex + 1;
END_WHILE
END_METHOD

(****************************************************************************************************<br>
© Syntegon Group.<br>
All rights reserved, also regarding any disposal, exploitation, reproduction, editing, distribution,<br>
as well as in the event of applications for industrial property rights.<br>
*****************************************************************************************************<br>
DESCRIPTION:<br>
A program value: node vi_dn_Parent is the parent of node vi_dn_Node (m_Link in role 0). Idempotent: call it every<br>
cycle after the declaration, before m_Cycle.<br>
*****************************************************************************************************<br>
OUTPUT VALUES:<br>
FALSE as m_Link.<br>
****************************************************************************************************)
METHOD m_SetParent : BOOL
VAR_INPUT
	vi_dn_Node							: DINT;	// [-] id of the child
	vi_dn_Parent						: DINT;	// [-] id of its parent
END_VAR
m_SetParent := m_Link(vi_dn_Node := vi_dn_Node, vi_un_Role := 0, vi_dn_Target := vi_dn_Parent);
END_METHOD

(****************************************************************************************************<br>
© Syntegon Group.<br>
All rights reserved, also regarding any disposal, exploitation, reproduction, editing, distribution,<br>
as well as in the event of applications for industrial property rights.<br>
*****************************************************************************************************<br>
DESCRIPTION:<br>
Makes the declared node vi_dn_Node the root node: the one node without a parent, from which every node in use<br>
hangs. Idempotent: call it every cycle after m_DeclareNode. A topology has one root node: another one is refused.<br>
*****************************************************************************************************<br>
OUTPUT VALUES:<br>
FALSE for a node not declared, or a second root node.<br>
****************************************************************************************************)
METHOD m_SetRoot : BOOL
VAR_INPUT
	vi_dn_Node							: DINT;	// [-] the node's id
END_VAR
m_SetRoot := m_NodeIndex(vi_dn_Id := vi_dn_Node) >= 0
	AND (vo_Config.nRootNode = 0 OR vo_Config.nRootNode = vi_dn_Node);
IF m_SetRoot THEN
	vo_Config.nRootNode := vi_dn_Node;
END_IF
END_METHOD

END_FUNCTION_BLOCK

// ---- POUs/_FC_GetVersionSynConfig.TcPOU
(****************************************************************************************************<br>
© Syntegon Group.<br>
All rights reserved, also regarding any disposal, exploitation, reproduction, editing, distribution,<br>
as well as in the event of applications for industrial property rights.<br>
*****************************************************************************************************<br>
DESCRIPTION:<br>
Runtime-readable version of the Syn_Config library.<br>
*****************************************************************************************************<br>
VERSION         ¦ DATE       ¦ NAME      ¦ CHANGE<br>
Syn_Config 1.0.0 ¦ 2026-11-10 ¦ J.Willner ¦ Parameter sets of conveyors and Deltas (ADR 0017, protocol 1)<br>
Syn_Config 1.1.0 ¦ 2026-11-10 ¦ J.Willner ¦ Every other component type (#24)<br>
Syn_Config 2.0.0 ¦ 2026-11-11 ¦ J.Willner ¦ Gripper fingers in the robots' sets (protocol 2, #25)<br>
Syn_Config 2.0.1 ¦ 2026-11-12 ¦ J.Willner ¦ SynVisu as a placeholder: the application chooses its version<br>
Syn_Config 2.1.0 ¦ 2026-11-14 ¦ J.Willner ¦ Machine FB: recipe fields and machine commands (protocol 3, #43)<br>
Syn_Config 2.2.0 ¦ 2026-11-14 ¦ J.Willner ¦ Recipe fields: label, description, visibility condition (protocol 4, #49)<br>
Syn_Config 2.3.0 ¦ 2026-11-14 ¦ J.Willner ¦ One staging lifecycle; m_PassOn passes the pose on (Syn_Visu 10.0.0)<br>
Syn_Config 2.4.0 ¦ 2026-11-19 ¦ J.Willner ¦ Topology FB: nodes, roles and program links (protocol 5, #56)<br>
****************************************************************************************************)
FUNCTION _FC_GetVersionSynConfig : UINT
VAR_INPUT
	vi_n_VersionElement					: INT;	// [-] 1 = major, 2 = minor, 3 = revision
END_VAR

CASE vi_n_VersionElement OF
	1: _FC_GetVersionSynConfig := 2;
	2: _FC_GetVersionSynConfig := 4;
	3: _FC_GetVersionSynConfig := 0;
ELSE
	_FC_GetVersionSynConfig := 16#FFFF;
END_CASE

END_FUNCTION

// ---- POUs/_FB_ConfigBodyComponent.TcPOU
(****************************************************************************************************<br>
© Syntegon Group.<br>
All rights reserved, also regarding any disposal, exploitation, reproduction, editing, distribution,<br>
as well as in the event of applications for industrial property rights.<br>
*****************************************************************************************************<br>
DESCRIPTION:<br>
Base of the parameter FBs of components drawn from their bodies (_FB_ConfigVision, _FB_ConfigSensor,<br>
_FB_ConfigStation, ADR 0017): their pose, origin shift and zones, written by the configurator, taken over when<br>
the application allows it. The bodies are hardware and stay the application's. Typical cycle:<br>
  fb_VisionParam.m_Register(vio_Manifest := GVL_Config.stManifest, vi_udn_Id := fb_Vision.m_Id());<br>
  fb_VisionParam.m_Cycle(vio_Default := VisionDefault, vio_Set := VisionSet, vi_b_ApplyAllowed := b_Stopped);<br>
  fb_Vision.m_Configure(vi_lr_FieldLength := 400, ...);<br>
  fb_VisionParam.m_PassOn(vio_Visu := fb_Vision);<br>
Not used directly.<br>
*****************************************************************************************************<br>
OUTPUT VALUES:<br>
vo_Config is the contract structure the gateway reads and writes at the path in the config manifest.<br>
*****************************************************************************************************<br>
VERSION         ¦ DATE       ¦ NAME      ¦ CHANGE<br>
Syn_Config 1.1.0 ¦ 2026-11-10 ¦ J.Willner ¦ New<br>
Syn_Config 2.3.0 ¦ 2026-11-14 ¦ J.Willner ¦ m_Cycle through m_HandleStaging; m_PassOnBody passes the pose on<br>
****************************************************************************************************)
FUNCTION_BLOCK ABSTRACT _FB_ConfigBodyComponent EXTENDS _FB_ConfigComponent
VAR_OUTPUT
	vo_Config							: ST_ConfigBodyComponent;	// contract structure of the gateway
END_VAR

(****************************************************************************************************<br>
© Syntegon Group.<br>
All rights reserved, also regarding any disposal, exploitation, reproduction, editing, distribution,<br>
as well as in the event of applications for industrial property rights.<br>
*****************************************************************************************************<br>
DESCRIPTION:<br>
All effective values (zones, ...), for the application's own logic.<br>
****************************************************************************************************)
METHOD m_Active : ST_ConfigBodyComponentParam
m_Active := vo_Config.stActive;
END_METHOD

(****************************************************************************************************<br>
© Syntegon Group.<br>
All rights reserved, also regarding any disposal, exploitation, reproduction, editing, distribution,<br>
as well as in the event of applications for industrial property rights.<br>
*****************************************************************************************************<br>
DESCRIPTION:<br>
Every cycle: handles a staged set or a reset (a set only while vi_b_ApplyAllowed), keeps the active set in<br>
vio_Set and gives the effective values in vo_Config.stActive: the active set while one is valid, else the<br>
program values vio_Default.<br>
*****************************************************************************************************<br>
OUTPUT VALUES:<br>
TRUE in the cycle a set was taken over or reset.<br>
****************************************************************************************************)
METHOD m_Cycle : BOOL
VAR_IN_OUT CONSTANT
	vio_Default							: ST_ConfigBodyComponentParam;	// the application's program values
END_VAR
VAR_IN_OUT
	vio_Set								: ST_ConfigBodyComponentSet;	// the application's VAR PERSISTENT active set
END_VAR
VAR_INPUT
	vi_b_ApplyAllowed					: BOOL;	// [-] a staged set may be taken over now, e.g. while the machine stands
END_VAR
VAR
	b_TempTakeOver						: BOOL;	// the staged set was taken over: copy it
END_VAR
m_Cycle := m_HandleStaging(vio_Staging := vo_Config.stStaging, vio_Status := vo_Config.stStatus, vio_b_Valid := vio_Set.bValid,
	vio_udn_Version := vio_Set.nVersion, vio_udn_LastVersion := vio_Set.nLastVersion, vi_b_ApplyAllowed := vi_b_ApplyAllowed,
	vo_b_TakeOver => b_TempTakeOver);
IF b_TempTakeOver THEN
	vio_Set.stParam := vo_Config.stStaged;
END_IF


(****************************************************************************************************
EFFECTIVE VALUES
****************************************************************************************************)
IF vio_Set.bValid THEN
	vo_Config.stActive := vio_Set.stParam;
ELSE
	vo_Config.stActive := vio_Default;
END_IF
END_METHOD

(****************************************************************************************************<br>
© Syntegon Group.<br>
All rights reserved, also regarding any disposal, exploitation, reproduction, editing, distribution,<br>
as well as in the event of applications for industrial property rights.<br>
*****************************************************************************************************<br>
DESCRIPTION:<br>
Why a staged set cannot be taken over; '' when it can: more zones than the list holds or a zone on no conveyor<br>
(id 0).<br>
****************************************************************************************************)
METHOD PROTECTED m_InvalidStaged : STRING(80)
m_InvalidStaged := m_InvalidZones(vio_aZones := vo_Config.stStaged.aZones, vi_un_Count := vo_Config.stStaged.nZoneCount);
END_METHOD

